(* IEC 61131-3 sources: plc-st-coding-agent/progress/evidence/f14_v10_full_20261113/jobs/codex_deepseek-v4pro, 82 files *)

(* ---- public-easy-01.candidate_01.st ---- *)
FUNCTION_BLOCK AutomatedFillingLineControl
(* ENGINEERING_CONTRACT
Stage0 idle: all outputs OFF; bottleSensor activates Pump_Motor (PUB001).
Pump_Motor: holds until cleaningConfirm; off by cleaningConfirm (PUB002).
Filling_Valve: set by cleaningConfirm; holds until fillingConfirm; off by fillingConfirm (PUB003).
Capping_Machine: set by fillingConfirm; holds until cappingConfirm; off by cappingConfirm (PUB004).
Packing_Machine: set by cappingConfirm; holds until packingConfirm; off by packingConfirm (PUB005).
Completion_Light: set by packingConfirm; holds until finishedButton; off by finishedButton (PUB006).
Same-scan priority: process only current stage trigger; at most one stage advance per scan.
Units/boundaries: BOOL outputs, integer stage 0..5; no timer or delay used.
*)
(* CONTRACT_RULES [
{"kind":"hold_until_reset","output":"Pump_Motor","set_input":"bottleSensor","reset_input":"cleaningConfirmButton"},
{"kind":"hold_until_reset","output":"Filling_Valve","set_input":"cleaningConfirmButton","reset_input":"fillingConfirmButton"},
{"kind":"hold_until_reset","output":"Capping_Machine","set_input":"fillingConfirmButton","reset_input":"cappingConfirmButton"},
{"kind":"hold_until_reset","output":"Packing_Machine","set_input":"cappingConfirmButton","reset_input":"packingConfirmButton"},
{"kind":"hold_until_reset","output":"Completion_Light","set_input":"packingConfirmButton","reset_input":"finishedButton"}
] *)
VAR_INPUT
    bottleSensor : BOOL;
    cleaningConfirmButton : BOOL;
    fillingConfirmButton : BOOL;
    cappingConfirmButton : BOOL;
    packingConfirmButton : BOOL;
    finishedButton : BOOL;
END_VAR
VAR_OUTPUT
    Pump_Motor : BOOL;
    Filling_Valve : BOOL;
    Capping_Machine : BOOL;
    Packing_Machine : BOOL;
    Completion_Light : BOOL;
END_VAR
VAR
    tmp_Stage : INT := 0;
END_VAR

IF tmp_Stage = 0 THEN
    IF bottleSensor THEN
        tmp_Stage := 1;
    END_IF;
ELSIF tmp_Stage = 1 THEN
    IF cleaningConfirmButton THEN
        tmp_Stage := 2;
    END_IF;
ELSIF tmp_Stage = 2 THEN
    IF fillingConfirmButton THEN
        tmp_Stage := 3;
    END_IF;
ELSIF tmp_Stage = 3 THEN
    IF cappingConfirmButton THEN
        tmp_Stage := 4;
    END_IF;
ELSIF tmp_Stage = 4 THEN
    IF packingConfirmButton THEN
        tmp_Stage := 5;
    END_IF;
ELSIF tmp_Stage = 5 THEN
    IF finishedButton THEN
        tmp_Stage := 0;
    END_IF;
END_IF;

Pump_Motor := (tmp_Stage = 1);
Filling_Valve := (tmp_Stage = 2);
Capping_Machine := (tmp_Stage = 3);
Packing_Machine := (tmp_Stage = 4);
Completion_Light := (tmp_Stage = 5);

END_FUNCTION_BLOCK

(* ---- public-easy-01.candidate_02.st ---- *)
FUNCTION_BLOCK AutomatedFillingLineControl
(* ENGINEERING_CONTRACT
Stage0 idle: all outputs OFF; bottleSensor activates Pump_Motor (PUB001).
Pump_Motor: holds until cleaningConfirm; off by cleaningConfirm (PUB002).
Filling_Valve: set by cleaningConfirm; holds until fillingConfirm; off by fillingConfirm (PUB003).
Capping_Machine: set by fillingConfirm; holds until cappingConfirm; off by cappingConfirm (PUB004).
Packing_Machine: set by cappingConfirm; holds until packingConfirm; off by packingConfirm (PUB005).
Completion_Light: set by packingConfirm; holds until finishedButton; off by finishedButton (PUB006).
Same-scan priority: process only current stage trigger; at most one stage advance per scan.
Units/boundaries: BOOL outputs, integer stage 0..5; no timer or delay used.
*)
(* CONTRACT_RULES [] *)
VAR_INPUT
    bottleSensor : BOOL;
    cleaningConfirmButton : BOOL;
    fillingConfirmButton : BOOL;
    cappingConfirmButton : BOOL;
    packingConfirmButton : BOOL;
    finishedButton : BOOL;
END_VAR
VAR_OUTPUT
    Pump_Motor : BOOL;
    Filling_Valve : BOOL;
    Capping_Machine : BOOL;
    Packing_Machine : BOOL;
    Completion_Light : BOOL;
END_VAR
VAR
    tmp_Stage : INT := 0;
END_VAR

IF tmp_Stage = 0 THEN
    IF bottleSensor THEN
        tmp_Stage := 1;
    END_IF;
ELSIF tmp_Stage = 1 THEN
    IF cleaningConfirmButton THEN
        tmp_Stage := 2;
    END_IF;
ELSIF tmp_Stage = 2 THEN
    IF fillingConfirmButton THEN
        tmp_Stage := 3;
    END_IF;
ELSIF tmp_Stage = 3 THEN
    IF cappingConfirmButton THEN
        tmp_Stage := 4;
    END_IF;
ELSIF tmp_Stage = 4 THEN
    IF packingConfirmButton THEN
        tmp_Stage := 5;
    END_IF;
ELSIF tmp_Stage = 5 THEN
    IF finishedButton THEN
        tmp_Stage := 0;
    END_IF;
END_IF;

Pump_Motor := (tmp_Stage = 1);
Filling_Valve := (tmp_Stage = 2);
Capping_Machine := (tmp_Stage = 3);
Packing_Machine := (tmp_Stage = 4);
Completion_Light := (tmp_Stage = 5);

END_FUNCTION_BLOCK

(* ---- public-easy-01.raw_candidate_01.st ---- *)
FUNCTION_BLOCK AutomatedFillingLineControl
(* ENGINEERING_CONTRACT
Stage0 idle: all outputs OFF; bottleSensor activates Pump_Motor (PUB001).
Pump_Motor: holds until cleaningConfirm; off by cleaningConfirm (PUB002).
Filling_Valve: set by cleaningConfirm; holds until fillingConfirm; off by fillingConfirm (PUB003).
Capping_Machine: set by fillingConfirm; holds until cappingConfirm; off by cappingConfirm (PUB004).
Packing_Machine: set by cappingConfirm; holds until packingConfirm; off by packingConfirm (PUB005).
Completion_Light: set by packingConfirm; holds until finishedButton; off by finishedButton (PUB006).
Same-scan priority: process only current stage trigger; at most one stage advance per scan.
Units/boundaries: BOOL outputs, integer stage 0..5; no timer or delay used.
*)
(* CONTRACT_RULES [
{"kind":"hold_until_reset","output":"Pump_Motor","set_input":"bottleSensor","reset_input":"cleaningConfirmButton"},
{"kind":"hold_until_reset","output":"Filling_Valve","set_input":"cleaningConfirmButton","reset_input":"fillingConfirmButton"},
{"kind":"hold_until_reset","output":"Capping_Machine","set_input":"fillingConfirmButton","reset_input":"cappingConfirmButton"},
{"kind":"hold_until_reset","output":"Packing_Machine","set_input":"cappingConfirmButton","reset_input":"packingConfirmButton"},
{"kind":"hold_until_reset","output":"Completion_Light","set_input":"packingConfirmButton","reset_input":"finishedButton"}
] *)
VAR_INPUT
    bottleSensor : BOOL;
    cleaningConfirmButton : BOOL;
    fillingConfirmButton : BOOL;
    cappingConfirmButton : BOOL;
    packingConfirmButton : BOOL;
    finishedButton : BOOL;
END_VAR
VAR_OUTPUT
    Pump_Motor : BOOL;
    Filling_Valve : BOOL;
    Capping_Machine : BOOL;
    Packing_Machine : BOOL;
    Completion_Light : BOOL;
END_VAR
VAR
    tmp_Stage : INT := 0;
END_VAR

IF tmp_Stage = 0 THEN
    IF bottleSensor THEN
        tmp_Stage := 1;
    END_IF;
ELSIF tmp_Stage = 1 THEN
    IF cleaningConfirmButton THEN
        tmp_Stage := 2;
    END_IF;
ELSIF tmp_Stage = 2 THEN
    IF fillingConfirmButton THEN
        tmp_Stage := 3;
    END_IF;
ELSIF tmp_Stage = 3 THEN
    IF cappingConfirmButton THEN
        tmp_Stage := 4;
    END_IF;
ELSIF tmp_Stage = 4 THEN
    IF packingConfirmButton THEN
        tmp_Stage := 5;
    END_IF;
ELSIF tmp_Stage = 5 THEN
    IF finishedButton THEN
        tmp_Stage := 0;
    END_IF;
END_IF;

Pump_Motor := (tmp_Stage = 1);
Filling_Valve := (tmp_Stage = 2);
Capping_Machine := (tmp_Stage = 3);
Packing_Machine := (tmp_Stage = 4);
Completion_Light := (tmp_Stage = 5);

END_FUNCTION_BLOCK

(* ---- public-easy-01.raw_candidate_02.st ---- *)
FUNCTION_BLOCK AutomatedFillingLineControl
(* ENGINEERING_CONTRACT
Stage0 idle: all outputs OFF; bottleSensor activates Pump_Motor (PUB001).
Pump_Motor: holds until cleaningConfirm; off by cleaningConfirm (PUB002).
Filling_Valve: set by cleaningConfirm; holds until fillingConfirm; off by fillingConfirm (PUB003).
Capping_Machine: set by fillingConfirm; holds until cappingConfirm; off by cappingConfirm (PUB004).
Packing_Machine: set by cappingConfirm; holds until packingConfirm; off by packingConfirm (PUB005).
Completion_Light: set by packingConfirm; holds until finishedButton; off by finishedButton (PUB006).
Same-scan priority: process only current stage trigger; at most one stage advance per scan.
Units/boundaries: BOOL outputs, integer stage 0..5; no timer or delay used.
*)
(* CONTRACT_RULES [] *)
VAR_INPUT
    bottleSensor : BOOL;
    cleaningConfirmButton : BOOL;
    fillingConfirmButton : BOOL;
    cappingConfirmButton : BOOL;
    packingConfirmButton : BOOL;
    finishedButton : BOOL;
END_VAR
VAR_OUTPUT
    Pump_Motor : BOOL;
    Filling_Valve : BOOL;
    Capping_Machine : BOOL;
    Packing_Machine : BOOL;
    Completion_Light : BOOL;
END_VAR
VAR
    tmp_Stage : INT := 0;
END_VAR

IF tmp_Stage = 0 THEN
    IF bottleSensor THEN
        tmp_Stage := 1;
    END_IF;
ELSIF tmp_Stage = 1 THEN
    IF cleaningConfirmButton THEN
        tmp_Stage := 2;
    END_IF;
ELSIF tmp_Stage = 2 THEN
    IF fillingConfirmButton THEN
        tmp_Stage := 3;
    END_IF;
ELSIF tmp_Stage = 3 THEN
    IF cappingConfirmButton THEN
        tmp_Stage := 4;
    END_IF;
ELSIF tmp_Stage = 4 THEN
    IF packingConfirmButton THEN
        tmp_Stage := 5;
    END_IF;
ELSIF tmp_Stage = 5 THEN
    IF finishedButton THEN
        tmp_Stage := 0;
    END_IF;
END_IF;

Pump_Motor := (tmp_Stage = 1);
Filling_Valve := (tmp_Stage = 2);
Capping_Machine := (tmp_Stage = 3);
Packing_Machine := (tmp_Stage = 4);
Completion_Light := (tmp_Stage = 5);

END_FUNCTION_BLOCK

(* ---- public-easy-02.candidate_01.st ---- *)
FUNCTION_BLOCK FB
(* ENGINEERING_CONTRACT
- PUB001: per-cycle edge detection on all 32 bits of DWORD value.
- hasChanged: on when current value <> retained lastValue; off otherwise.
- risingBits[i]: on when lastValue[i]=0 and value[i]=1; noOfRisingBits counts bits 0..31.
- hasRisingEdges: on when noOfRisingBits > 0; off otherwise.
- fallingBits[i]: on when lastValue[i]=1 and value[i]=0; noOfFallingBits counts bits 0..31.
- hasFallingEdges: on when noOfFallingBits > 0; off otherwise.
- Retention: only lastValue is retained. Outputs are recomputed every scan; no user reset.
- First-scan baseline: lastValue=0; unspecified, tested consistently with previous value zero.
- Priority: compare against old lastValue first, then store current value at scan end.
- Bounds: counts are USINT 0..32; masks cover DWORD bits 0..31.
*)
(* CONTRACT_RULES [] *)
VAR_INPUT
    value : DWORD;
END_VAR
VAR_OUTPUT
    hasChanged : BOOL;
    hasRisingEdges : BOOL;
    risingBits : DWORD;
    noOfRisingBits : USINT;
    hasFallingEdges : BOOL;
    fallingBits : DWORD;
    noOfFallingBits : USINT;
END_VAR
VAR
    lastValue : DWORD;
    tmp_rising : DWORD;
    tmp_falling : DWORD;
    tmp_i : INT;
END_VAR

tmp_rising := (NOT lastValue) AND value;
tmp_falling := lastValue AND (NOT value);

hasChanged := value <> lastValue;
risingBits := tmp_rising;
fallingBits := tmp_falling;

noOfRisingBits := 0;
noOfFallingBits := 0;

FOR tmp_i := 0 TO 31 DO
    IF (tmp_rising AND SHL(DWORD#1, tmp_i)) <> DWORD#0 THEN
        noOfRisingBits := noOfRisingBits + 1;
    END_IF;
    IF (tmp_falling AND SHL(DWORD#1, tmp_i)) <> DWORD#0 THEN
        noOfFallingBits := noOfFallingBits + 1;
    END_IF;
END_FOR;

hasRisingEdges := noOfRisingBits > 0;
hasFallingEdges := noOfFallingBits > 0;

lastValue := value;
END_FUNCTION_BLOCK

(* ---- public-easy-02.raw_candidate_01.st ---- *)
FUNCTION_BLOCK FB
(* ENGINEERING_CONTRACT
- PUB001: per-cycle edge detection on all 32 bits of DWORD value.
- hasChanged: on when current value <> retained lastValue; off otherwise.
- risingBits[i]: on when lastValue[i]=0 and value[i]=1; noOfRisingBits counts bits 0..31.
- hasRisingEdges: on when noOfRisingBits > 0; off otherwise.
- fallingBits[i]: on when lastValue[i]=1 and value[i]=0; noOfFallingBits counts bits 0..31.
- hasFallingEdges: on when noOfFallingBits > 0; off otherwise.
- Retention: only lastValue is retained. Outputs are recomputed every scan; no user reset.
- First-scan baseline: lastValue=0; unspecified, tested consistently with previous value zero.
- Priority: compare against old lastValue first, then store current value at scan end.
- Bounds: counts are USINT 0..32; masks cover DWORD bits 0..31.
*)
(* CONTRACT_RULES [] *)
VAR_INPUT
    value : DWORD;
END_VAR
VAR_OUTPUT
    hasChanged : BOOL;
    hasRisingEdges : BOOL;
    risingBits : DWORD;
    noOfRisingBits : USINT;
    hasFallingEdges : BOOL;
    fallingBits : DWORD;
    noOfFallingBits : USINT;
END_VAR
VAR
    lastValue : DWORD;
    tmp_rising : DWORD;
    tmp_falling : DWORD;
    tmp_i : INT;
END_VAR

tmp_rising := (NOT lastValue) AND value;
tmp_falling := lastValue AND (NOT value);

hasChanged := value <> lastValue;
risingBits := tmp_rising;
fallingBits := tmp_falling;

noOfRisingBits := 0;
noOfFallingBits := 0;

FOR tmp_i := 0 TO 31 DO
    IF (tmp_rising AND SHL(DWORD#1, tmp_i)) <> DWORD#0 THEN
        noOfRisingBits := noOfRisingBits + 1;
    END_IF;
    IF (tmp_falling AND SHL(DWORD#1, tmp_i)) <> DWORD#0 THEN
        noOfFallingBits := noOfFallingBits + 1;
    END_IF;
END_FOR;

hasRisingEdges := noOfRisingBits > 0;
hasFallingEdges := noOfFallingBits > 0;

lastValue := value;
END_FUNCTION_BLOCK

(* ---- public-easy-03.candidate_01.st ---- *)
FUNCTION_BLOCK AlarmHandling
(* ENGINEERING_CONTRACT
  hiAlarm (PUB001): activate only when Value > hiLevel; hold across deadband until deactivation.
  hiAlarm deactivation (PUB001): deactivate only when Value < hiLevel - hystWindow (strict).
  loAlarm (PUB001): activate only when Value < loLevel; hold across deadband until deactivation.
  loAlarm deactivation (PUB001): deactivate only when Value > loLevel + hystWindow (strict).
  error/status (PUB006, PUB007): normal scan sets error:=FALSE and status:=0.
  Same-scan priority: loLevel >= hiLevel (16#8001) is checked first and invokes RETURN before alarm evaluation.
  hystWindow >= hiLevel - loLevel (16#8002) is checked next and suppresses normal alarm evaluation via ELSE.
  Retention: alarm outputs persist while inside their respective hysteresis deadband.
  Units: REAL values are dimensionless; status is a hexadecimal WORD code.
  Unspecified: behavior for NaN/Inf, negative hystWindow, and historical alarm state during error scans.
*)
(* CONTRACT_RULES [] *)
VAR_INPUT
    Value      : REAL;
    hiLevel    : REAL;
    loLevel    : REAL;
    hystWindow : REAL;
END_VAR
VAR_OUTPUT
    hiAlarm : BOOL;
    loAlarm : BOOL;
    error   : BOOL;
    status  : WORD;
END_VAR
VAR
END_VAR

    error := FALSE;
    status := 0;

    IF loLevel >= hiLevel THEN
        error := TRUE;
        status := WORD#16#8001;
        RETURN;
    END_IF;

    IF hystWindow >= (hiLevel - loLevel) THEN
        error := TRUE;
        status := WORD#16#8002;
    ELSE
        IF Value > hiLevel THEN
            hiAlarm := TRUE;
        ELSIF Value < (hiLevel - hystWindow) THEN
            hiAlarm := FALSE;
        END_IF;

        IF Value < loLevel THEN
            loAlarm := TRUE;
        ELSIF Value > (loLevel + hystWindow) THEN
            loAlarm := FALSE;
        END_IF;
    END_IF;

END_FUNCTION_BLOCK

(* ---- public-easy-03.raw_candidate_01.st ---- *)
FUNCTION_BLOCK AlarmHandling
(* ENGINEERING_CONTRACT
  hiAlarm (PUB001): activate only when Value > hiLevel; hold across deadband until deactivation.
  hiAlarm deactivation (PUB001): deactivate only when Value < hiLevel - hystWindow (strict).
  loAlarm (PUB001): activate only when Value < loLevel; hold across deadband until deactivation.
  loAlarm deactivation (PUB001): deactivate only when Value > loLevel + hystWindow (strict).
  error/status (PUB006, PUB007): normal scan sets error:=FALSE and status:=0.
  Same-scan priority: loLevel >= hiLevel (16#8001) is checked first and invokes RETURN before alarm evaluation.
  hystWindow >= hiLevel - loLevel (16#8002) is checked next and suppresses normal alarm evaluation via ELSE.
  Retention: alarm outputs persist while inside their respective hysteresis deadband.
  Units: REAL values are dimensionless; status is a hexadecimal WORD code.
  Unspecified: behavior for NaN/Inf, negative hystWindow, and historical alarm state during error scans.
*)
(* CONTRACT_RULES [] *)
VAR_INPUT
    Value      : REAL;
    hiLevel    : REAL;
    loLevel    : REAL;
    hystWindow : REAL;
END_VAR
VAR_OUTPUT
    hiAlarm : BOOL;
    loAlarm : BOOL;
    error   : BOOL;
    status  : WORD;
END_VAR
VAR
END_VAR

    error := FALSE;
    status := 0;

    IF loLevel >= hiLevel THEN
        error := TRUE;
        status := WORD#16#8001;
        RETURN;
    END_IF;

    IF hystWindow >= (hiLevel - loLevel) THEN
        error := TRUE;
        status := WORD#16#8002;
    ELSE
        IF Value > hiLevel THEN
            hiAlarm := TRUE;
        ELSIF Value < (hiLevel - hystWindow) THEN
            hiAlarm := FALSE;
        END_IF;

        IF Value < loLevel THEN
            loAlarm := TRUE;
        ELSIF Value > (loLevel + hystWindow) THEN
            loAlarm := FALSE;
        END_IF;
    END_IF;

END_FUNCTION_BLOCK

(* ---- public-easy-04.candidate_01.st ---- *)
FUNCTION_BLOCK JamPumpControl
VAR_INPUT
    VISCOSITY_OK : BOOL;
    PASTE_E_STOP_NC : BOOL;
    DebounceTime : TIME;
    CycleTime : TIME;
END_VAR
VAR_OUTPUT
    VFD_RUN : BOOL := FALSE;
    PUMP_MAINT_DUE : BOOL := FALSE;
    PUMP_RUNTIME_ACC : LTIME := LTIME#0s;
END_VAR
VAR
    viscosityValid : BOOL := FALSE;
    viscosityDebounce : TON;
END_VAR

(* ENGINEERING_CONTRACT
Viscosity state PUB001/PUB002: activation after VISCOSITY_OK remains TRUE for DebounceTime via TON; invalidated immediately on VISCOSITY_OK FALSE; already-valid state retained through E-stop; incomplete debounce timing cleared on E-stop FALSE.
VFD_RUN PUB002/PUB005: activation = PASTE_E_STOP_NC AND viscosityValid; no hold/latch; E-stop FALSE disables run immediately in same scan; initialized FALSE.
PUMP_RUNTIME_ACC PUB003/PUB005: activation after current VFD_RUN computation; adds TIME_TO_LTIME(CycleTime) while VFD_RUN TRUE; retained while stopped; no explicit reset; initialized LTIME#0s.
PUMP_MAINT_DUE PUB004/PUB005: activation and retention when PUMP_RUNTIME_ACC >= LTIME#500h; no reset; informational only, never gates run/permissive; initialized FALSE.
Same-scan priority: E-stop disable and viscosity invalidation occur before run accumulation; maintenance computation is independent.
Units/boundaries: DebounceTime TIME ms, CycleTime TIME ms, PUMP_RUNTIME_ACC LTIME ns, maintenance threshold >= 500 h.
*)

(* CONTRACT_RULES [] *)

viscosityDebounce(IN := VISCOSITY_OK AND PASTE_E_STOP_NC,
                  PT := DebounceTime);

IF NOT VISCOSITY_OK THEN
    viscosityValid := FALSE;
ELSIF viscosityDebounce.Q THEN
    viscosityValid := TRUE;
END_IF;

VFD_RUN := PASTE_E_STOP_NC AND viscosityValid;

IF VFD_RUN THEN
    PUMP_RUNTIME_ACC := PUMP_RUNTIME_ACC + TIME_TO_LTIME(CycleTime);
END_IF;

IF PUMP_RUNTIME_ACC >= LTIME#500h THEN
    PUMP_MAINT_DUE := TRUE;
END_IF;

END_FUNCTION_BLOCK

(* ---- public-easy-04.raw_candidate_01.st ---- *)
FUNCTION_BLOCK JamPumpControl
VAR_INPUT
    VISCOSITY_OK : BOOL;
    PASTE_E_STOP_NC : BOOL;
    DebounceTime : TIME;
    CycleTime : TIME;
END_VAR
VAR_OUTPUT
    VFD_RUN : BOOL := FALSE;
    PUMP_MAINT_DUE : BOOL := FALSE;
    PUMP_RUNTIME_ACC : LTIME := LTIME#0s;
END_VAR
VAR
    viscosityValid : BOOL := FALSE;
    viscosityDebounce : TON;
END_VAR

(* ENGINEERING_CONTRACT
Viscosity state PUB001/PUB002: activation after VISCOSITY_OK remains TRUE for DebounceTime via TON; invalidated immediately on VISCOSITY_OK FALSE; already-valid state retained through E-stop; incomplete debounce timing cleared on E-stop FALSE.
VFD_RUN PUB002/PUB005: activation = PASTE_E_STOP_NC AND viscosityValid; no hold/latch; E-stop FALSE disables run immediately in same scan; initialized FALSE.
PUMP_RUNTIME_ACC PUB003/PUB005: activation after current VFD_RUN computation; adds TIME_TO_LTIME(CycleTime) while VFD_RUN TRUE; retained while stopped; no explicit reset; initialized LTIME#0s.
PUMP_MAINT_DUE PUB004/PUB005: activation and retention when PUMP_RUNTIME_ACC >= LTIME#500h; no reset; informational only, never gates run/permissive; initialized FALSE.
Same-scan priority: E-stop disable and viscosity invalidation occur before run accumulation; maintenance computation is independent.
Units/boundaries: DebounceTime TIME ms, CycleTime TIME ms, PUMP_RUNTIME_ACC LTIME ns, maintenance threshold >= 500 h.
*)

(* CONTRACT_RULES [] *)

viscosityDebounce(IN := VISCOSITY_OK AND PASTE_E_STOP_NC,
                  PT := DebounceTime);

IF NOT VISCOSITY_OK THEN
    viscosityValid := FALSE;
ELSIF viscosityDebounce.Q THEN
    viscosityValid := TRUE;
END_IF;

VFD_RUN := PASTE_E_STOP_NC AND viscosityValid;

IF VFD_RUN THEN
    PUMP_RUNTIME_ACC := PUMP_RUNTIME_ACC + TIME_TO_LTIME(CycleTime);
END_IF;

IF PUMP_RUNTIME_ACC >= LTIME#500h THEN
    PUMP_MAINT_DUE := TRUE;
END_IF;

END_FUNCTION_BLOCK

(* ---- public-easy-05.candidate_01.st ---- *)
FUNCTION_BLOCK WeldGapAlarmFB
VAR_INPUT
    Gap_Exceeded        : BOOL;
    Weld_E_Stop_NC      : BOOL;
    DebounceTime        : TIME;
END_VAR
VAR_OUTPUT
    Operator_Alert       : BOOL;
    Weld_Soft_Start_Active : BOOL;
END_VAR
VAR
    InitTimer       : TON;
    DebounceTimer   : TON;
    InitComplete    : BOOL;
    NormalMonitor   : BOOL;
END_VAR

(*
ENGINEERING_CONTRACT
- Operator_Alert: activates only when initialization is complete, E-stop is inactive,
  and Gap_Exceeded has remained TRUE for DebounceTime (PUB003, PUB004).
  It is FALSE during the 5 s initialization period (PUB002).
- Operator_Alert reset: immediately FALSE when Gap_Exceeded becomes FALSE or E-stop
  becomes active; normal-monitoring conditions must remain true to hold it (PUB003, PUB004).
- Debounce timing: accumulates only during initialized normal monitoring with E-stop
  inactive and resets when Gap_Exceeded is FALSE or E-stop is active (PUB002, PUB003, PUB004).
- Weld_Soft_Start_Active: TRUE only during the first 5 s after power-up, independent of
  E-stop state; it is not a speed ramp (PUB002, PUB005). E-stop state is not specified
  for this output.
- Boundaries/units: initialization is fixed T#5S; DebounceTime uses TIME milliseconds.
  TON activation occurs at elapsed time >= PT.
*)

InitTimer(IN := TRUE, PT := T#5S);
InitComplete := InitTimer.Q;
NormalMonitor := InitComplete AND Weld_E_Stop_NC;

DebounceTimer(IN := Gap_Exceeded AND NormalMonitor, PT := DebounceTime);

Operator_Alert := NormalMonitor AND DebounceTimer.Q;
Weld_Soft_Start_Active := NOT InitComplete;

(* CONTRACT_RULES [] *)
END_FUNCTION_BLOCK

(* ---- public-easy-05.raw_candidate_01.st ---- *)
FUNCTION_BLOCK WeldGapAlarmFB
VAR_INPUT
    Gap_Exceeded        : BOOL;
    Weld_E_Stop_NC      : BOOL;
    DebounceTime        : TIME;
END_VAR
VAR_OUTPUT
    Operator_Alert       : BOOL;
    Weld_Soft_Start_Active : BOOL;
END_VAR
VAR
    InitTimer       : TON;
    DebounceTimer   : TON;
    InitComplete    : BOOL;
    NormalMonitor   : BOOL;
END_VAR

(*
ENGINEERING_CONTRACT
- Operator_Alert: activates only when initialization is complete, E-stop is inactive,
  and Gap_Exceeded has remained TRUE for DebounceTime (PUB003, PUB004).
  It is FALSE during the 5 s initialization period (PUB002).
- Operator_Alert reset: immediately FALSE when Gap_Exceeded becomes FALSE or E-stop
  becomes active; normal-monitoring conditions must remain true to hold it (PUB003, PUB004).
- Debounce timing: accumulates only during initialized normal monitoring with E-stop
  inactive and resets when Gap_Exceeded is FALSE or E-stop is active (PUB002, PUB003, PUB004).
- Weld_Soft_Start_Active: TRUE only during the first 5 s after power-up, independent of
  E-stop state; it is not a speed ramp (PUB002, PUB005). E-stop state is not specified
  for this output.
- Boundaries/units: initialization is fixed T#5S; DebounceTime uses TIME milliseconds.
  TON activation occurs at elapsed time >= PT.
*)

InitTimer(IN := TRUE, PT := T#5S);
InitComplete := InitTimer.Q;
NormalMonitor := InitComplete AND Weld_E_Stop_NC;

DebounceTimer(IN := Gap_Exceeded AND NormalMonitor, PT := DebounceTime);

Operator_Alert := NormalMonitor AND DebounceTimer.Q;
Weld_Soft_Start_Active := NOT InitComplete;

(* CONTRACT_RULES [] *)
END_FUNCTION_BLOCK

(* ---- public-easy-06.candidate_01.st ---- *)
FUNCTION_BLOCK AerationBlowerDelayedStart
VAR_INPUT
    DO_LOW : BOOL;
    AERATION_E_STOP_NC : BOOL;
END_VAR
VAR_OUTPUT
    BLOWER_RUN : BOOL;
    AERATION_BLOWER_CYCLE_COUNT : UINT;
END_VAR
VAR
    tmp_StartDelay : TON;
    tmp_PrevRun : BOOL := FALSE;
END_VAR

(*
ENGINEERING_CONTRACT
- BLOWER_RUN activation: only when DO_LOW and AERATION_E_STOP_NC have both been TRUE for T#5s (PUB001).
- BLOWER_RUN retention/hold: remains TRUE only while both enabling conditions remain TRUE; no separate latch is used.
- BLOWER_RUN explicit reset/deactivation: any FALSE of DO_LOW or AERATION_E_STOP_NC clears timer IN immediately, so output and timing reset (PUB002).
- AERATION_BLOWER_CYCLE_COUNT activation: increments once on each BLOWER_RUN FALSE->TRUE transition; not repeated during continuous run (PUB003).
- AERATION_BLOWER_CYCLE_COUNT reset: initialized to zero at power-up; no task-specified runtime reset is implemented (PUB004).
- Same-scan priority: current DO_LOW/E_STOP condition directly gates TON.IN before timer Q and edge counting are evaluated.
- Units/boundaries: delay is 5 000 ms (T#5s); cycle count is UINT and unspecified at maximum rollover.
*)
(* CONTRACT_RULES [] *)

tmp_StartDelay(IN := DO_LOW AND AERATION_E_STOP_NC, PT := T#5S);

BLOWER_RUN := tmp_StartDelay.Q;

IF BLOWER_RUN AND NOT tmp_PrevRun THEN
    AERATION_BLOWER_CYCLE_COUNT := AERATION_BLOWER_CYCLE_COUNT + 1;
END_IF;

tmp_PrevRun := BLOWER_RUN;

END_FUNCTION_BLOCK

(* ---- public-easy-06.raw_candidate_01.st ---- *)
FUNCTION_BLOCK AerationBlowerDelayedStart
VAR_INPUT
    DO_LOW : BOOL;
    AERATION_E_STOP_NC : BOOL;
END_VAR
VAR_OUTPUT
    BLOWER_RUN : BOOL;
    AERATION_BLOWER_CYCLE_COUNT : UINT;
END_VAR
VAR
    tmp_StartDelay : TON;
    tmp_PrevRun : BOOL := FALSE;
END_VAR

(*
ENGINEERING_CONTRACT
- BLOWER_RUN activation: only when DO_LOW and AERATION_E_STOP_NC have both been TRUE for T#5s (PUB001).
- BLOWER_RUN retention/hold: remains TRUE only while both enabling conditions remain TRUE; no separate latch is used.
- BLOWER_RUN explicit reset/deactivation: any FALSE of DO_LOW or AERATION_E_STOP_NC clears timer IN immediately, so output and timing reset (PUB002).
- AERATION_BLOWER_CYCLE_COUNT activation: increments once on each BLOWER_RUN FALSE->TRUE transition; not repeated during continuous run (PUB003).
- AERATION_BLOWER_CYCLE_COUNT reset: initialized to zero at power-up; no task-specified runtime reset is implemented (PUB004).
- Same-scan priority: current DO_LOW/E_STOP condition directly gates TON.IN before timer Q and edge counting are evaluated.
- Units/boundaries: delay is 5 000 ms (T#5s); cycle count is UINT and unspecified at maximum rollover.
*)
(* CONTRACT_RULES [] *)

tmp_StartDelay(IN := DO_LOW AND AERATION_E_STOP_NC, PT := T#5S);

BLOWER_RUN := tmp_StartDelay.Q;

IF BLOWER_RUN AND NOT tmp_PrevRun THEN
    AERATION_BLOWER_CYCLE_COUNT := AERATION_BLOWER_CYCLE_COUNT + 1;
END_IF;

tmp_PrevRun := BLOWER_RUN;

END_FUNCTION_BLOCK

(* ---- public-hard-02.candidate_01.st ---- *)
FUNCTION_BLOCK FlexibleProcessingControl
(* ENGINEERING_CONTRACT
   conveyorLeft  : active while moving to a lower-numbered station; deactivates when the destination sensor is detected or when final delivery to station 5 is complete. No separate reset input is specified. Same-scan arrival clears both conveyors (PUB002/PUB003/PUB005).
   conveyorRight : active while moving to a higher-numbered station; deactivates when the destination sensor is detected or when final delivery to station 5 is complete. No separate reset input is specified. Same-scan arrival clears both conveyors (PUB002/PUB003/PUB005).
   Processing wait: retained in phase after arrival at station 2, 3, or 4. The matching completion input starts the next sequence movement in the same scan it is detected (PUB002/PUB003).
   Start condition: sensor1 AND station1Start initiates processing from processSequence[1]; after transition, START is not re-evaluated until the current product cycle is finished (PUB001/PUB006).
   Boundaries: processLength is active in the range 1..8; active sequence positions are processSequence[1] through processSequence[processLength]. Stations are compared as USINT values 1..5 (PUB004/PUB006).
*)
(* CONTRACT_RULES [] *)
VAR_INPUT
    processLength : USINT;
    sensor1 : BOOL;
    sensor2 : BOOL;
    sensor3 : BOOL;
    sensor4 : BOOL;
    sensor5 : BOOL;
    station1Start : BOOL;
    station2Complete : BOOL;
    station3Complete : BOOL;
    station4Complete : BOOL;
    processSequence : ARRAY[1..8] OF USINT;
END_VAR
VAR_OUTPUT
    conveyorLeft : BOOL;
    conveyorRight : BOOL;
END_VAR
VAR
    tmp_phase : USINT := 0;
    tmp_seqIndex : USINT := 1;
    tmp_currentStation : USINT := 1;
    tmp_targetStation : USINT := 0;
    tmp_destSensor : BOOL := FALSE;
    tmp_completeSignal : BOOL := FALSE;
    tmp_activeLength : USINT := 1;
END_VAR

tmp_activeLength := processLength;
IF tmp_activeLength > 8 THEN
    tmp_activeLength := 8;
END_IF;
IF tmp_activeLength < 1 THEN
    tmp_activeLength := 1;
END_IF;

conveyorLeft := FALSE;
conveyorRight := FALSE;

IF tmp_phase = 0 THEN
    IF sensor1 AND station1Start THEN
        tmp_seqIndex := 1;
        IF tmp_seqIndex <= tmp_activeLength THEN
            tmp_targetStation := processSequence[tmp_seqIndex];
            tmp_phase := 1;
        END_IF;
    END_IF;
END_IF;

IF tmp_phase = 2 THEN
    tmp_completeSignal := FALSE;
    CASE tmp_currentStation OF
        2:
            tmp_completeSignal := station2Complete;
        3:
            tmp_completeSignal := station3Complete;
        4:
            tmp_completeSignal := station4Complete;
    ELSE
        tmp_completeSignal := FALSE;
    END_CASE;

    IF tmp_completeSignal THEN
        IF tmp_seqIndex < tmp_activeLength THEN
            tmp_seqIndex := tmp_seqIndex + 1;
            IF tmp_seqIndex <= tmp_activeLength THEN
                tmp_targetStation := processSequence[tmp_seqIndex];
                tmp_phase := 1;
            END_IF;
        END_IF;
    END_IF;
END_IF;

IF tmp_phase = 1 THEN
    IF tmp_targetStation > tmp_currentStation THEN
        conveyorRight := TRUE;
    ELSIF tmp_targetStation < tmp_currentStation THEN
        conveyorLeft := TRUE;
    END_IF;

    tmp_destSensor := FALSE;
    CASE tmp_targetStation OF
        2:
            tmp_destSensor := sensor2;
        3:
            tmp_destSensor := sensor3;
        4:
            tmp_destSensor := sensor4;
        5:
            tmp_destSensor := sensor5;
    ELSE
        tmp_destSensor := FALSE;
    END_CASE;

    IF tmp_destSensor THEN
        conveyorLeft := FALSE;
        conveyorRight := FALSE;
        tmp_currentStation := tmp_targetStation;

        IF tmp_currentStation = 5 THEN
            tmp_phase := 3;
        ELSE
            tmp_phase := 2;
        END_IF;
    END_IF;
END_IF;

END_FUNCTION_BLOCK

(* ---- public-hard-02.candidate_02.st ---- *)
FUNCTION_BLOCK FlexibleProcessingControl
(* ENGINEERING_CONTRACT
   conveyorLeft  : active while moving to a lower-numbered station; deactivates when the destination sensor is detected or when final delivery to station 5 is complete. No separate reset input is specified. Same-scan arrival clears both conveyors (PUB002/PUB003/PUB005).
   conveyorRight : active while moving to a higher-numbered station; deactivates when the destination sensor is detected or when final delivery to station 5 is complete. No separate reset input is specified. Same-scan arrival clears both conveyors (PUB002/PUB003/PUB005).
   Processing wait: retained in phase after arrival at station 2, 3, or 4. The matching completion input starts the next sequence movement in the same scan it is detected (PUB002/PUB003).
   Start condition: sensor1 AND station1Start initiates processing from processSequence[1]; after transition, START is not re-evaluated until the current product cycle is finished (PUB001/PUB006). On a new start, current station returns to 1.
   Boundaries: processLength is active in the range 1..8; active sequence positions are processSequence[1] through processSequence[processLength]. Stations are compared as USINT values 1..5 (PUB004/PUB006).
*)
(* CONTRACT_RULES [] *)
VAR_INPUT
    processLength : USINT;
    sensor1 : BOOL;
    sensor2 : BOOL;
    sensor3 : BOOL;
    sensor4 : BOOL;
    sensor5 : BOOL;
    station1Start : BOOL;
    station2Complete : BOOL;
    station3Complete : BOOL;
    station4Complete : BOOL;
    processSequence : ARRAY[1..8] OF USINT;
END_VAR
VAR_OUTPUT
    conveyorLeft : BOOL;
    conveyorRight : BOOL;
END_VAR
VAR
    tmp_phase : USINT := 0;
    tmp_seqIndex : USINT := 1;
    tmp_currentStation : USINT := 1;
    tmp_targetStation : USINT := 0;
    tmp_destSensor : BOOL := FALSE;
    tmp_completeSignal : BOOL := FALSE;
    tmp_activeLength : USINT := 1;
END_VAR

tmp_activeLength := processLength;
IF tmp_activeLength > 8 THEN
    tmp_activeLength := 8;
END_IF;
IF tmp_activeLength < 1 THEN
    tmp_activeLength := 1;
END_IF;

conveyorLeft := FALSE;
conveyorRight := FALSE;

IF tmp_phase = 0 THEN
    IF sensor1 AND station1Start THEN
        tmp_seqIndex := 1;
        tmp_currentStation := 1;
        IF tmp_seqIndex <= tmp_activeLength THEN
            tmp_targetStation := processSequence[tmp_seqIndex];
            tmp_phase := 1;
        END_IF;
    END_IF;
END_IF;

IF tmp_phase = 2 THEN
    tmp_completeSignal := FALSE;
    CASE tmp_currentStation OF
        2:
            tmp_completeSignal := station2Complete;
        3:
            tmp_completeSignal := station3Complete;
        4:
            tmp_completeSignal := station4Complete;
    ELSE
        tmp_completeSignal := FALSE;
    END_CASE;

    IF tmp_completeSignal THEN
        IF tmp_seqIndex < tmp_activeLength THEN
            tmp_seqIndex := tmp_seqIndex + 1;
            IF tmp_seqIndex <= tmp_activeLength THEN
                tmp_targetStation := processSequence[tmp_seqIndex];
                tmp_phase := 1;
            END_IF;
        END_IF;
    END_IF;
END_IF;

IF tmp_phase = 1 THEN
    IF tmp_targetStation > tmp_currentStation THEN
        conveyorRight := TRUE;
    ELSIF tmp_targetStation < tmp_currentStation THEN
        conveyorLeft := TRUE;
    END_IF;

    tmp_destSensor := FALSE;
    CASE tmp_targetStation OF
        2:
            tmp_destSensor := sensor2;
        3:
            tmp_destSensor := sensor3;
        4:
            tmp_destSensor := sensor4;
        5:
            tmp_destSensor := sensor5;
    ELSE
        tmp_destSensor := FALSE;
    END_CASE;

    IF tmp_destSensor THEN
        conveyorLeft := FALSE;
        conveyorRight := FALSE;
        tmp_currentStation := tmp_targetStation;

        IF tmp_currentStation = 5 THEN
            tmp_phase := 0;
        ELSE
            tmp_phase := 2;
        END_IF;
    END_IF;
END_IF;

END_FUNCTION_BLOCK

(* ---- public-hard-02.raw_candidate_01.st ---- *)
FUNCTION_BLOCK FlexibleProcessingControl
(* ENGINEERING_CONTRACT
   conveyorLeft  : active while moving to a lower-numbered station; deactivates when the destination sensor is detected or when final delivery to station 5 is complete. No separate reset input is specified. Same-scan arrival clears both conveyors (PUB002/PUB003/PUB005).
   conveyorRight : active while moving to a higher-numbered station; deactivates when the destination sensor is detected or when final delivery to station 5 is complete. No separate reset input is specified. Same-scan arrival clears both conveyors (PUB002/PUB003/PUB005).
   Processing wait: retained in phase after arrival at station 2, 3, or 4. The matching completion input starts the next sequence movement in the same scan it is detected (PUB002/PUB003).
   Start condition: sensor1 AND station1Start initiates processing from processSequence[1]; after transition, START is not re-evaluated until the current product cycle is finished (PUB001/PUB006).
   Boundaries: processLength is active in the range 1..8; active sequence positions are processSequence[1] through processSequence[processLength]. Stations are compared as USINT values 1..5 (PUB004/PUB006).
*)
(* CONTRACT_RULES [] *)
VAR_INPUT
    processLength : USINT;
    sensor1 : BOOL;
    sensor2 : BOOL;
    sensor3 : BOOL;
    sensor4 : BOOL;
    sensor5 : BOOL;
    station1Start : BOOL;
    station2Complete : BOOL;
    station3Complete : BOOL;
    station4Complete : BOOL;
    processSequence : ARRAY[1..8] OF USINT;
END_VAR
VAR_OUTPUT
    conveyorLeft : BOOL;
    conveyorRight : BOOL;
END_VAR
VAR
    tmp_phase : USINT := 0;
    tmp_seqIndex : USINT := 1;
    tmp_currentStation : USINT := 1;
    tmp_targetStation : USINT := 0;
    tmp_destSensor : BOOL := FALSE;
    tmp_completeSignal : BOOL := FALSE;
    tmp_activeLength : USINT := 1;
END_VAR

tmp_activeLength := processLength;
IF tmp_activeLength > 8 THEN
    tmp_activeLength := 8;
END_IF;
IF tmp_activeLength < 1 THEN
    tmp_activeLength := 1;
END_IF;

conveyorLeft := FALSE;
conveyorRight := FALSE;

IF tmp_phase = 0 THEN
    IF sensor1 AND station1Start THEN
        tmp_seqIndex := 1;
        IF tmp_seqIndex <= tmp_activeLength THEN
            tmp_targetStation := processSequence[tmp_seqIndex];
            tmp_phase := 1;
        END_IF;
    END_IF;
END_IF;

IF tmp_phase = 2 THEN
    tmp_completeSignal := FALSE;
    CASE tmp_currentStation OF
        2:
            tmp_completeSignal := station2Complete;
        3:
            tmp_completeSignal := station3Complete;
        4:
            tmp_completeSignal := station4Complete;
    ELSE
        tmp_completeSignal := FALSE;
    END_CASE;

    IF tmp_completeSignal THEN
        IF tmp_seqIndex < tmp_activeLength THEN
            tmp_seqIndex := tmp_seqIndex + 1;
            IF tmp_seqIndex <= tmp_activeLength THEN
                tmp_targetStation := processSequence[tmp_seqIndex];
                tmp_phase := 1;
            END_IF;
        END_IF;
    END_IF;
END_IF;

IF tmp_phase = 1 THEN
    IF tmp_targetStation > tmp_currentStation THEN
        conveyorRight := TRUE;
    ELSIF tmp_targetStation < tmp_currentStation THEN
        conveyorLeft := TRUE;
    END_IF;

    tmp_destSensor := FALSE;
    CASE tmp_targetStation OF
        2:
            tmp_destSensor := sensor2;
        3:
            tmp_destSensor := sensor3;
        4:
            tmp_destSensor := sensor4;
        5:
            tmp_destSensor := sensor5;
    ELSE
        tmp_destSensor := FALSE;
    END_CASE;

    IF tmp_destSensor THEN
        conveyorLeft := FALSE;
        conveyorRight := FALSE;
        tmp_currentStation := tmp_targetStation;

        IF tmp_currentStation = 5 THEN
            tmp_phase := 3;
        ELSE
            tmp_phase := 2;
        END_IF;
    END_IF;
END_IF;

END_FUNCTION_BLOCK

(* ---- public-hard-02.raw_candidate_02.st ---- *)
FUNCTION_BLOCK FlexibleProcessingControl
(* ENGINEERING_CONTRACT
   conveyorLeft  : active while moving to a lower-numbered station; deactivates when the destination sensor is detected or when final delivery to station 5 is complete. No separate reset input is specified. Same-scan arrival clears both conveyors (PUB002/PUB003/PUB005).
   conveyorRight : active while moving to a higher-numbered station; deactivates when the destination sensor is detected or when final delivery to station 5 is complete. No separate reset input is specified. Same-scan arrival clears both conveyors (PUB002/PUB003/PUB005).
   Processing wait: retained in phase after arrival at station 2, 3, or 4. The matching completion input starts the next sequence movement in the same scan it is detected (PUB002/PUB003).
   Start condition: sensor1 AND station1Start initiates processing from processSequence[1]; after transition, START is not re-evaluated until the current product cycle is finished (PUB001/PUB006). On a new start, current station returns to 1.
   Boundaries: processLength is active in the range 1..8; active sequence positions are processSequence[1] through processSequence[processLength]. Stations are compared as USINT values 1..5 (PUB004/PUB006).
*)
(* CONTRACT_RULES [] *)
VAR_INPUT
    processLength : USINT;
    sensor1 : BOOL;
    sensor2 : BOOL;
    sensor3 : BOOL;
    sensor4 : BOOL;
    sensor5 : BOOL;
    station1Start : BOOL;
    station2Complete : BOOL;
    station3Complete : BOOL;
    station4Complete : BOOL;
    processSequence : ARRAY[1..8] OF USINT;
END_VAR
VAR_OUTPUT
    conveyorLeft : BOOL;
    conveyorRight : BOOL;
END_VAR
VAR
    tmp_phase : USINT := 0;
    tmp_seqIndex : USINT := 1;
    tmp_currentStation : USINT := 1;
    tmp_targetStation : USINT := 0;
    tmp_destSensor : BOOL := FALSE;
    tmp_completeSignal : BOOL := FALSE;
    tmp_activeLength : USINT := 1;
END_VAR

tmp_activeLength := processLength;
IF tmp_activeLength > 8 THEN
    tmp_activeLength := 8;
END_IF;
IF tmp_activeLength < 1 THEN
    tmp_activeLength := 1;
END_IF;

conveyorLeft := FALSE;
conveyorRight := FALSE;

IF tmp_phase = 0 THEN
    IF sensor1 AND station1Start THEN
        tmp_seqIndex := 1;
        tmp_currentStation := 1;
        IF tmp_seqIndex <= tmp_activeLength THEN
            tmp_targetStation := processSequence[tmp_seqIndex];
            tmp_phase := 1;
        END_IF;
    END_IF;
END_IF;

IF tmp_phase = 2 THEN
    tmp_completeSignal := FALSE;
    CASE tmp_currentStation OF
        2:
            tmp_completeSignal := station2Complete;
        3:
            tmp_completeSignal := station3Complete;
        4:
            tmp_completeSignal := station4Complete;
    ELSE
        tmp_completeSignal := FALSE;
    END_CASE;

    IF tmp_completeSignal THEN
        IF tmp_seqIndex < tmp_activeLength THEN
            tmp_seqIndex := tmp_seqIndex + 1;
            IF tmp_seqIndex <= tmp_activeLength THEN
                tmp_targetStation := processSequence[tmp_seqIndex];
                tmp_phase := 1;
            END_IF;
        END_IF;
    END_IF;
END_IF;

IF tmp_phase = 1 THEN
    IF tmp_targetStation > tmp_currentStation THEN
        conveyorRight := TRUE;
    ELSIF tmp_targetStation < tmp_currentStation THEN
        conveyorLeft := TRUE;
    END_IF;

    tmp_destSensor := FALSE;
    CASE tmp_targetStation OF
        2:
            tmp_destSensor := sensor2;
        3:
            tmp_destSensor := sensor3;
        4:
            tmp_destSensor := sensor4;
        5:
            tmp_destSensor := sensor5;
    ELSE
        tmp_destSensor := FALSE;
    END_CASE;

    IF tmp_destSensor THEN
        conveyorLeft := FALSE;
        conveyorRight := FALSE;
        tmp_currentStation := tmp_targetStation;

        IF tmp_currentStation = 5 THEN
            tmp_phase := 0;
        ELSE
            tmp_phase := 2;
        END_IF;
    END_IF;
END_IF;

END_FUNCTION_BLOCK

(* ---- public-hard-03.candidate_01.st ---- *)
TYPE ST_Recipe :
STRUCT
    recipeID : INT;
    ingredientType : INT;
    ingredientRatio : REAL;
    productionTemperature : REAL;
END_STRUCT
END_TYPE;

(* ENGINEERING_CONTRACT
   Outputs: success flags are same-scan level, not latched; they deactivate on the next scan (PUB003-PUB005).
   recipeQueryResult: updated only for a successful query; otherwise zeroed each scan (PUB002).
   error/status: cleared at scan start; first operation error in the scan retains error and code (PUB002-PUB005).
   Add: duplicate check before empty-slot check; uses first empty index; whole struct copy (PUB003).
   Delete: nonzero-ID match; sets only recipeID to 0 (PUB004).
   Modify: nonzero-ID match; whole struct replacement (PUB005).
   Query: nonzero-ID match; whole struct copy to result; missing ID gives 16#8001 (PUB002).
   Array bounds: 1..10; recipeID=0 denotes unused slot and is never returned as a stored recipe.
   Multiple requests: unspecified; processed add/delete/modify/query in interface order on evolving database.
*)
(* CONTRACT_RULES [] *)

FUNCTION_BLOCK RecipeManagementSystem
VAR_INPUT
    addRecipe : BOOL;
    deleteRecipe : BOOL;
    modifyRecipe : BOOL;
    queryRecipe : BOOL;
    recipeIn : ST_Recipe;
END_VAR
VAR_OUTPUT
    recipeAdded : BOOL;
    recipeDeleted : BOOL;
    recipeModified : BOOL;
    recipeQueryResult : ST_Recipe;
    error : BOOL;
    status : WORD;
END_VAR
VAR_IN_OUT
    recipe : ARRAY[1..10] OF ST_Recipe;
END_VAR
VAR
    tmp_i : INT;
    tmp_foundIndex : INT;
    tmp_emptyIndex : INT;
    tmp_found : BOOL;
END_VAR

recipeAdded := FALSE;
recipeDeleted := FALSE;
recipeModified := FALSE;
recipeQueryResult.recipeID := 0;
recipeQueryResult.ingredientType := 0;
recipeQueryResult.ingredientRatio := 0.0;
recipeQueryResult.productionTemperature := 0.0;
error := FALSE;
status := 16#0000;

IF addRecipe THEN
    tmp_found := FALSE;
    tmp_emptyIndex := 0;

    FOR tmp_i := 1 TO 10 DO
        IF recipe[tmp_i].recipeID = recipeIn.recipeID THEN
            tmp_found := TRUE;
        END_IF;

        IF (recipe[tmp_i].recipeID = 0) AND (tmp_emptyIndex = 0) THEN
            tmp_emptyIndex := tmp_i;
        END_IF;
    END_FOR;

    IF tmp_found THEN
        IF NOT error THEN
            error := TRUE;
            status := 16#8002;
        END_IF;
    ELSIF tmp_emptyIndex = 0 THEN
        IF NOT error THEN
            error := TRUE;
            status := 16#8003;
        END_IF;
    ELSE
        recipe[tmp_emptyIndex] := recipeIn;
        recipeAdded := TRUE;
    END_IF;
END_IF;

IF deleteRecipe THEN
    tmp_found := FALSE;
    tmp_foundIndex := 0;

    FOR tmp_i := 1 TO 10 DO
        IF (recipe[tmp_i].recipeID <> 0) AND
           (recipe[tmp_i].recipeID = recipeIn.recipeID) THEN
            tmp_found := TRUE;
            tmp_foundIndex := tmp_i;
        END_IF;
    END_FOR;

    IF NOT tmp_found THEN
        IF NOT error THEN
            error := TRUE;
            status := 16#8004;
        END_IF;
    ELSE
        recipe[tmp_foundIndex].recipeID := 0;
        recipeDeleted := TRUE;
    END_IF;
END_IF;

IF modifyRecipe THEN
    tmp_found := FALSE;
    tmp_foundIndex := 0;

    FOR tmp_i := 1 TO 10 DO
        IF (recipe[tmp_i].recipeID <> 0) AND
           (recipe[tmp_i].recipeID = recipeIn.recipeID) THEN
            tmp_found := TRUE;
            tmp_foundIndex := tmp_i;
        END_IF;
    END_FOR;

    IF NOT tmp_found THEN
        IF NOT error THEN
            error := TRUE;
            status := 16#8005;
        END_IF;
    ELSE
        recipe[tmp_foundIndex] := recipeIn;
        recipeModified := TRUE;
    END_IF;
END_IF;

IF queryRecipe THEN
    tmp_found := FALSE;
    tmp_foundIndex := 0;

    FOR tmp_i := 1 TO 10 DO
        IF (recipe[tmp_i].recipeID <> 0) AND
           (recipe[tmp_i].recipeID = recipeIn.recipeID) THEN
            tmp_found := TRUE;
            tmp_foundIndex := tmp_i;
        END_IF;
    END_FOR;

    IF NOT tmp_found THEN
        IF NOT error THEN
            error := TRUE;
            status := 16#8001;
        END_IF;
    ELSE
        recipeQueryResult := recipe[tmp_foundIndex];
    END_IF;
END_IF;

END_FUNCTION_BLOCK

(* ---- public-hard-03.candidate_02.st ---- *)
TYPE ST_Recipe :
STRUCT
    recipeID : INT;
    ingredientType : INT;
    ingredientRatio : REAL;
    productionTemperature : REAL;
END_STRUCT
END_TYPE;

(* ENGINEERING_CONTRACT
   Outputs: success flags are same-scan level, not latched; they deactivate on the next scan (PUB003-PUB005).
   recipeQueryResult: updated only for a successful query; otherwise zeroed each scan (PUB002).
   error/status: cleared at scan start; a reported operation error retains error and code for that invocation (PUB002-PUB005).
   Add: duplicate check before empty-slot check; uses first empty index; whole struct copy (PUB003).
   Delete: nonzero-ID match; sets only recipeID to 0 (PUB004).
   Modify: nonzero-ID match; whole struct replacement (PUB005).
   Query: nonzero-ID match; whole struct copy to result; missing ID gives 16#8001 (PUB002).
   Array bounds: 1..10; recipeID=0 denotes unused slot and is never returned as a stored recipe.
   Multiple requests: unspecified by the public contract. They are reported as an unsupported combination with
   error=TRUE, status=16#8000, no database update, no success flag, and no query result.
*)
(* CONTRACT_RULES [] *)

FUNCTION_BLOCK RecipeManagementSystem
VAR_INPUT
    addRecipe : BOOL;
    deleteRecipe : BOOL;
    modifyRecipe : BOOL;
    queryRecipe : BOOL;
    recipeIn : ST_Recipe;
END_VAR
VAR_OUTPUT
    recipeAdded : BOOL;
    recipeDeleted : BOOL;
    recipeModified : BOOL;
    recipeQueryResult : ST_Recipe;
    error : BOOL;
    status : WORD;
END_VAR
VAR_IN_OUT
    recipe : ARRAY[1..10] OF ST_Recipe;
END_VAR
VAR
    tmp_i : INT;
    tmp_foundIndex : INT;
    tmp_emptyIndex : INT;
    tmp_found : BOOL;
    tmp_cmdCount : INT;
END_VAR

recipeAdded := FALSE;
recipeDeleted := FALSE;
recipeModified := FALSE;
recipeQueryResult.recipeID := 0;
recipeQueryResult.ingredientType := 0;
recipeQueryResult.ingredientRatio := 0.0;
recipeQueryResult.productionTemperature := 0.0;
error := FALSE;
status := 16#0000;

tmp_cmdCount := 0;
IF addRecipe THEN
    tmp_cmdCount := tmp_cmdCount + 1;
END_IF;
IF deleteRecipe THEN
    tmp_cmdCount := tmp_cmdCount + 1;
END_IF;
IF modifyRecipe THEN
    tmp_cmdCount := tmp_cmdCount + 1;
END_IF;
IF queryRecipe THEN
    tmp_cmdCount := tmp_cmdCount + 1;
END_IF;

IF tmp_cmdCount > 1 THEN
    error := TRUE;
    status := 16#8000;
ELSE
    IF addRecipe THEN
        tmp_found := FALSE;
        tmp_emptyIndex := 0;

        FOR tmp_i := 1 TO 10 DO
            IF recipe[tmp_i].recipeID = recipeIn.recipeID THEN
                tmp_found := TRUE;
            END_IF;

            IF (recipe[tmp_i].recipeID = 0) AND (tmp_emptyIndex = 0) THEN
                tmp_emptyIndex := tmp_i;
            END_IF;
        END_FOR;

        IF tmp_found THEN
            IF NOT error THEN
                error := TRUE;
                status := 16#8002;
            END_IF;
        ELSIF tmp_emptyIndex = 0 THEN
            IF NOT error THEN
                error := TRUE;
                status := 16#8003;
            END_IF;
        ELSE
            recipe[tmp_emptyIndex] := recipeIn;
            recipeAdded := TRUE;
        END_IF;
    END_IF;

    IF deleteRecipe THEN
        tmp_found := FALSE;
        tmp_foundIndex := 0;

        FOR tmp_i := 1 TO 10 DO
            IF (recipe[tmp_i].recipeID <> 0) AND
               (recipe[tmp_i].recipeID = recipeIn.recipeID) THEN
                tmp_found := TRUE;
                tmp_foundIndex := tmp_i;
            END_IF;
        END_FOR;

        IF NOT tmp_found THEN
            IF NOT error THEN
                error := TRUE;
                status := 16#8004;
            END_IF;
        ELSE
            recipe[tmp_foundIndex].recipeID := 0;
            recipeDeleted := TRUE;
        END_IF;
    END_IF;

    IF modifyRecipe THEN
        tmp_found := FALSE;
        tmp_foundIndex := 0;

        FOR tmp_i := 1 TO 10 DO
            IF (recipe[tmp_i].recipeID <> 0) AND
               (recipe[tmp_i].recipeID = recipeIn.recipeID) THEN
                tmp_found := TRUE;
                tmp_foundIndex := tmp_i;
            END_IF;
        END_FOR;

        IF NOT tmp_found THEN
            IF NOT error THEN
                error := TRUE;
                status := 16#8005;
            END_IF;
        ELSE
            recipe[tmp_foundIndex] := recipeIn;
            recipeModified := TRUE;
        END_IF;
    END_IF;

    IF queryRecipe THEN
        tmp_found := FALSE;
        tmp_foundIndex := 0;

        FOR tmp_i := 1 TO 10 DO
            IF (recipe[tmp_i].recipeID <> 0) AND
               (recipe[tmp_i].recipeID = recipeIn.recipeID) THEN
                tmp_found := TRUE;
                tmp_foundIndex := tmp_i;
            END_IF;
        END_FOR;

        IF NOT tmp_found THEN
            IF NOT error THEN
                error := TRUE;
                status := 16#8001;
            END_IF;
        ELSE
            recipeQueryResult := recipe[tmp_foundIndex];
        END_IF;
    END_IF;
END_IF;

END_FUNCTION_BLOCK

(* ---- public-hard-03.raw_candidate_01.st ---- *)
TYPE ST_Recipe :
STRUCT
    recipeID : INT;
    ingredientType : INT;
    ingredientRatio : REAL;
    productionTemperature : REAL;
END_STRUCT
END_TYPE

(* ENGINEERING_CONTRACT
   Outputs: success flags are same-scan level, not latched; they deactivate on the next scan (PUB003-PUB005).
   recipeQueryResult: updated only for a successful query; otherwise zeroed each scan (PUB002).
   error/status: cleared at scan start; first operation error in the scan retains error and code (PUB002-PUB005).
   Add: duplicate check before empty-slot check; uses first empty index; whole struct copy (PUB003).
   Delete: nonzero-ID match; sets only recipeID to 0 (PUB004).
   Modify: nonzero-ID match; whole struct replacement (PUB005).
   Query: nonzero-ID match; whole struct copy to result; missing ID gives 16#8001 (PUB002).
   Array bounds: 1..10; recipeID=0 denotes unused slot and is never returned as a stored recipe.
   Multiple requests: unspecified; processed add/delete/modify/query in interface order on evolving database.
*)
(* CONTRACT_RULES [] *)

FUNCTION_BLOCK RecipeManagementSystem
VAR_INPUT
    addRecipe : BOOL;
    deleteRecipe : BOOL;
    modifyRecipe : BOOL;
    queryRecipe : BOOL;
    recipeIn : ST_Recipe;
END_VAR
VAR_OUTPUT
    recipeAdded : BOOL;
    recipeDeleted : BOOL;
    recipeModified : BOOL;
    recipeQueryResult : ST_Recipe;
    error : BOOL;
    status : WORD;
END_VAR
VAR_IN_OUT
    recipe : ARRAY[1..10] OF ST_Recipe;
END_VAR
VAR
    tmp_i : INT;
    tmp_foundIndex : INT;
    tmp_emptyIndex : INT;
    tmp_found : BOOL;
END_VAR

recipeAdded := FALSE;
recipeDeleted := FALSE;
recipeModified := FALSE;
recipeQueryResult.recipeID := 0;
recipeQueryResult.ingredientType := 0;
recipeQueryResult.ingredientRatio := 0.0;
recipeQueryResult.productionTemperature := 0.0;
error := FALSE;
status := 16#0000;

IF addRecipe THEN
    tmp_found := FALSE;
    tmp_emptyIndex := 0;

    FOR tmp_i := 1 TO 10 DO
        IF recipe[tmp_i].recipeID = recipeIn.recipeID THEN
            tmp_found := TRUE;
        END_IF;

        IF (recipe[tmp_i].recipeID = 0) AND (tmp_emptyIndex = 0) THEN
            tmp_emptyIndex := tmp_i;
        END_IF;
    END_FOR;

    IF tmp_found THEN
        IF NOT error THEN
            error := TRUE;
            status := 16#8002;
        END_IF;
    ELSIF tmp_emptyIndex = 0 THEN
        IF NOT error THEN
            error := TRUE;
            status := 16#8003;
        END_IF;
    ELSE
        recipe[tmp_emptyIndex] := recipeIn;
        recipeAdded := TRUE;
    END_IF;
END_IF;

IF deleteRecipe THEN
    tmp_found := FALSE;
    tmp_foundIndex := 0;

    FOR tmp_i := 1 TO 10 DO
        IF (recipe[tmp_i].recipeID <> 0) AND
           (recipe[tmp_i].recipeID = recipeIn.recipeID) THEN
            tmp_found := TRUE;
            tmp_foundIndex := tmp_i;
        END_IF;
    END_FOR;

    IF NOT tmp_found THEN
        IF NOT error THEN
            error := TRUE;
            status := 16#8004;
        END_IF;
    ELSE
        recipe[tmp_foundIndex].recipeID := 0;
        recipeDeleted := TRUE;
    END_IF;
END_IF;

IF modifyRecipe THEN
    tmp_found := FALSE;
    tmp_foundIndex := 0;

    FOR tmp_i := 1 TO 10 DO
        IF (recipe[tmp_i].recipeID <> 0) AND
           (recipe[tmp_i].recipeID = recipeIn.recipeID) THEN
            tmp_found := TRUE;
            tmp_foundIndex := tmp_i;
        END_IF;
    END_FOR;

    IF NOT tmp_found THEN
        IF NOT error THEN
            error := TRUE;
            status := 16#8005;
        END_IF;
    ELSE
        recipe[tmp_foundIndex] := recipeIn;
        recipeModified := TRUE;
    END_IF;
END_IF;

IF queryRecipe THEN
    tmp_found := FALSE;
    tmp_foundIndex := 0;

    FOR tmp_i := 1 TO 10 DO
        IF (recipe[tmp_i].recipeID <> 0) AND
           (recipe[tmp_i].recipeID = recipeIn.recipeID) THEN
            tmp_found := TRUE;
            tmp_foundIndex := tmp_i;
        END_IF;
    END_FOR;

    IF NOT tmp_found THEN
        IF NOT error THEN
            error := TRUE;
            status := 16#8001;
        END_IF;
    ELSE
        recipeQueryResult := recipe[tmp_foundIndex];
    END_IF;
END_IF;

END_FUNCTION_BLOCK

(* ---- public-hard-03.raw_candidate_02.st ---- *)
TYPE ST_Recipe :
STRUCT
    recipeID : INT;
    ingredientType : INT;
    ingredientRatio : REAL;
    productionTemperature : REAL;
END_STRUCT
END_TYPE;

(* ENGINEERING_CONTRACT
   Outputs: success flags are same-scan level, not latched; they deactivate on the next scan (PUB003-PUB005).
   recipeQueryResult: updated only for a successful query; otherwise zeroed each scan (PUB002).
   error/status: cleared at scan start; a reported operation error retains error and code for that invocation (PUB002-PUB005).
   Add: duplicate check before empty-slot check; uses first empty index; whole struct copy (PUB003).
   Delete: nonzero-ID match; sets only recipeID to 0 (PUB004).
   Modify: nonzero-ID match; whole struct replacement (PUB005).
   Query: nonzero-ID match; whole struct copy to result; missing ID gives 16#8001 (PUB002).
   Array bounds: 1..10; recipeID=0 denotes unused slot and is never returned as a stored recipe.
   Multiple requests: unspecified by the public contract. They are reported as an unsupported combination with
   error=TRUE, status=16#8000, no database update, no success flag, and no query result.
*)
(* CONTRACT_RULES [] *)

FUNCTION_BLOCK RecipeManagementSystem
VAR_INPUT
    addRecipe : BOOL;
    deleteRecipe : BOOL;
    modifyRecipe : BOOL;
    queryRecipe : BOOL;
    recipeIn : ST_Recipe;
END_VAR
VAR_OUTPUT
    recipeAdded : BOOL;
    recipeDeleted : BOOL;
    recipeModified : BOOL;
    recipeQueryResult : ST_Recipe;
    error : BOOL;
    status : WORD;
END_VAR
VAR_IN_OUT
    recipe : ARRAY[1..10] OF ST_Recipe;
END_VAR
VAR
    tmp_i : INT;
    tmp_foundIndex : INT;
    tmp_emptyIndex : INT;
    tmp_found : BOOL;
    tmp_cmdCount : INT;
END_VAR

recipeAdded := FALSE;
recipeDeleted := FALSE;
recipeModified := FALSE;
recipeQueryResult.recipeID := 0;
recipeQueryResult.ingredientType := 0;
recipeQueryResult.ingredientRatio := 0.0;
recipeQueryResult.productionTemperature := 0.0;
error := FALSE;
status := 16#0000;

tmp_cmdCount := 0;
IF addRecipe THEN
    tmp_cmdCount := tmp_cmdCount + 1;
END_IF;
IF deleteRecipe THEN
    tmp_cmdCount := tmp_cmdCount + 1;
END_IF;
IF modifyRecipe THEN
    tmp_cmdCount := tmp_cmdCount + 1;
END_IF;
IF queryRecipe THEN
    tmp_cmdCount := tmp_cmdCount + 1;
END_IF;

IF tmp_cmdCount > 1 THEN
    error := TRUE;
    status := 16#8000;
ELSE
    IF addRecipe THEN
        tmp_found := FALSE;
        tmp_emptyIndex := 0;

        FOR tmp_i := 1 TO 10 DO
            IF recipe[tmp_i].recipeID = recipeIn.recipeID THEN
                tmp_found := TRUE;
            END_IF;

            IF (recipe[tmp_i].recipeID = 0) AND (tmp_emptyIndex = 0) THEN
                tmp_emptyIndex := tmp_i;
            END_IF;
        END_FOR;

        IF tmp_found THEN
            IF NOT error THEN
                error := TRUE;
                status := 16#8002;
            END_IF;
        ELSIF tmp_emptyIndex = 0 THEN
            IF NOT error THEN
                error := TRUE;
                status := 16#8003;
            END_IF;
        ELSE
            recipe[tmp_emptyIndex] := recipeIn;
            recipeAdded := TRUE;
        END_IF;
    END_IF;

    IF deleteRecipe THEN
        tmp_found := FALSE;
        tmp_foundIndex := 0;

        FOR tmp_i := 1 TO 10 DO
            IF (recipe[tmp_i].recipeID <> 0) AND
               (recipe[tmp_i].recipeID = recipeIn.recipeID) THEN
                tmp_found := TRUE;
                tmp_foundIndex := tmp_i;
            END_IF;
        END_FOR;

        IF NOT tmp_found THEN
            IF NOT error THEN
                error := TRUE;
                status := 16#8004;
            END_IF;
        ELSE
            recipe[tmp_foundIndex].recipeID := 0;
            recipeDeleted := TRUE;
        END_IF;
    END_IF;

    IF modifyRecipe THEN
        tmp_found := FALSE;
        tmp_foundIndex := 0;

        FOR tmp_i := 1 TO 10 DO
            IF (recipe[tmp_i].recipeID <> 0) AND
               (recipe[tmp_i].recipeID = recipeIn.recipeID) THEN
                tmp_found := TRUE;
                tmp_foundIndex := tmp_i;
            END_IF;
        END_FOR;

        IF NOT tmp_found THEN
            IF NOT error THEN
                error := TRUE;
                status := 16#8005;
            END_IF;
        ELSE
            recipe[tmp_foundIndex] := recipeIn;
            recipeModified := TRUE;
        END_IF;
    END_IF;

    IF queryRecipe THEN
        tmp_found := FALSE;
        tmp_foundIndex := 0;

        FOR tmp_i := 1 TO 10 DO
            IF (recipe[tmp_i].recipeID <> 0) AND
               (recipe[tmp_i].recipeID = recipeIn.recipeID) THEN
                tmp_found := TRUE;
                tmp_foundIndex := tmp_i;
            END_IF;
        END_FOR;

        IF NOT tmp_found THEN
            IF NOT error THEN
                error := TRUE;
                status := 16#8001;
            END_IF;
        ELSE
            recipeQueryResult := recipe[tmp_foundIndex];
        END_IF;
    END_IF;
END_IF;

END_FUNCTION_BLOCK

(* ---- public-hard-04.candidate_01.st ---- *)
FUNCTION_BLOCK FB_FIFO
VAR_INPUT
    enqueue : BOOL;
    dequeue : BOOL;
    reset : BOOL;
END_VAR
VAR_OUTPUT
    elementCount : DINT;
    status : WORD;
END_VAR
VAR_IN_OUT
    item : VARIANT;
    buffer : VARIANT;
END_VAR
VAR
    localCapacity : DINT;
    localLower : DINT;
    localHead : DINT;
    localTail : DINT;
    localCount : DINT;
    localNext : DINT;
    localLastEnqueue : BOOL;
    localLastDequeue : BOOL;
    localRisingEnqueue : BOOL;
    localRisingDequeue : BOOL;
END_VAR

(* ENGINEERING_CONTRACT
   validCount: activated by successful enqueue/dequeue; reset to 0 by reset (PUB001/PUB003).
   elementCount: mirror of persistent validCount each scan; reset sets it to 0 (PUB003/PUB004).
   status: default 16#0000; 16#8001 empty dequeue reject; 16#8002 full enqueue reject (PUB005).
   head/tail: internal only, initialized to buffer lower bound, advanced circularly (PUB006).
   priority: reset is processed before all queue operations (PUB003).
   same scan: caller precondition forbids simultaneous edges; if both occur enqueue is handled first (PUB002).
   full condition: validCount = capacity; empty condition: validCount = 0 (PUB004).
   capacity: UPPER_BOUND(buffer,1)-LOWER_BOUND(buffer,1)+1; indices are DINT (PUB004/PUB006).
   rejected operations: item and queue are not modified (PUB005).
   units/bounds: elementCount DINT 0..capacity; status WORD; no unconditional public BOOL latch.
*)

(* CONTRACT_RULES [] *)

IF localCapacity = 0 THEN
    localLower := LOWER_BOUND(buffer, 1);
    localCapacity := UPPER_BOUND(buffer, 1) - localLower + 1;
    localHead := localLower;
    localTail := localLower;
    localCount := 0;
END_IF;

status := WORD#16#0000;

localRisingEnqueue := enqueue AND NOT localLastEnqueue;
localRisingDequeue := dequeue AND NOT localLastDequeue;

IF reset THEN
    localCount := 0;
    localHead := localLower;
    localTail := localLower;
ELSE
    IF localRisingEnqueue THEN
        IF localCount < localCapacity THEN
            buffer[localTail] := item;
            localNext := localTail - localLower + 1;
            IF localNext >= localCapacity THEN
                localNext := 0;
            END_IF;
            localTail := localLower + localNext;
            localCount := localCount + 1;
        ELSE
            status := WORD#16#8002;
        END_IF;
    END_IF;

    IF localRisingDequeue THEN
        IF localCount > 0 THEN
            item := buffer[localHead];
            localNext := localHead - localLower + 1;
            IF localNext >= localCapacity THEN
                localNext := 0;
            END_IF;
            localHead := localLower + localNext;
            localCount := localCount - 1;
        ELSE
            status := WORD#16#8001;
        END_IF;
    END_IF;
END_IF;

elementCount := localCount;

localLastEnqueue := enqueue;
localLastDequeue := dequeue;

END_FUNCTION_BLOCK

(* ---- public-hard-04.raw_candidate_01.st ---- *)
FUNCTION_BLOCK FB_FIFO
VAR_INPUT
    enqueue : BOOL;
    dequeue : BOOL;
    reset : BOOL;
END_VAR
VAR_OUTPUT
    elementCount : DINT;
    status : WORD;
END_VAR
VAR_IN_OUT
    item : VARIANT;
    buffer : VARIANT;
END_VAR
VAR
    localCapacity : DINT;
    localLower : DINT;
    localHead : DINT;
    localTail : DINT;
    localCount : DINT;
    localNext : DINT;
    localLastEnqueue : BOOL;
    localLastDequeue : BOOL;
    localRisingEnqueue : BOOL;
    localRisingDequeue : BOOL;
END_VAR

(* ENGINEERING_CONTRACT
   validCount: activated by successful enqueue/dequeue; reset to 0 by reset (PUB001/PUB003).
   elementCount: mirror of persistent validCount each scan; reset sets it to 0 (PUB003/PUB004).
   status: default 16#0000; 16#8001 empty dequeue reject; 16#8002 full enqueue reject (PUB005).
   head/tail: internal only, initialized to buffer lower bound, advanced circularly (PUB006).
   priority: reset is processed before all queue operations (PUB003).
   same scan: caller precondition forbids simultaneous edges; if both occur enqueue is handled first (PUB002).
   full condition: validCount = capacity; empty condition: validCount = 0 (PUB004).
   capacity: UPPER_BOUND(buffer,1)-LOWER_BOUND(buffer,1)+1; indices are DINT (PUB004/PUB006).
   rejected operations: item and queue are not modified (PUB005).
   units/bounds: elementCount DINT 0..capacity; status WORD; no unconditional public BOOL latch.
*)

(* CONTRACT_RULES [] *)

IF localCapacity = 0 THEN
    localLower := LOWER_BOUND(buffer, 1);
    localCapacity := UPPER_BOUND(buffer, 1) - localLower + 1;
    localHead := localLower;
    localTail := localLower;
    localCount := 0;
END_IF;

status := WORD#16#0000;

localRisingEnqueue := enqueue AND NOT localLastEnqueue;
localRisingDequeue := dequeue AND NOT localLastDequeue;

IF reset THEN
    localCount := 0;
    localHead := localLower;
    localTail := localLower;
ELSE
    IF localRisingEnqueue THEN
        IF localCount < localCapacity THEN
            buffer[localTail] := item;
            localNext := localTail - localLower + 1;
            IF localNext >= localCapacity THEN
                localNext := 0;
            END_IF;
            localTail := localLower + localNext;
            localCount := localCount + 1;
        ELSE
            status := WORD#16#8002;
        END_IF;
    END_IF;

    IF localRisingDequeue THEN
        IF localCount > 0 THEN
            item := buffer[localHead];
            localNext := localHead - localLower + 1;
            IF localNext >= localCapacity THEN
                localNext := 0;
            END_IF;
            localHead := localLower + localNext;
            localCount := localCount - 1;
        ELSE
            status := WORD#16#8001;
        END_IF;
    END_IF;
END_IF;

elementCount := localCount;

localLastEnqueue := enqueue;
localLastDequeue := dequeue;

END_FUNCTION_BLOCK

(* ---- public-medium-01.candidate_01.st ---- *)
TYPE ST_Pump :
STRUCT
    priority : INT;
    selection : BOOL;
    RunComd : BOOL;
END_STRUCT
END_TYPE;

FUNCTION_BLOCK FB_MultiPumpSwitchingControl
(* ENGINEERING_CONTRACT
   - mode=FALSE: manual mode; RunComd follows selection (PUB001/PUB002).
   - mode=TRUE: automatic mode; select three pumps with highest priority (PUB001/PUB003).
   - start: activates run enable; stop: deactivates run enable and stops all pumps (PUB002/PUB004).
   - Same-scan stop priority: if stop=TRUE, stop wins over start.
   - Run command is evaluated as selected AND run enable each scan.
   - Larger priority wins. Equal priority is unspecified; lower array index wins.
   - Mode transition with run enable retained is unspecified; retained run enable is used.
*)
(* CONTRACT_RULES [] *)
VAR
    runEnable : BOOL := FALSE;
    tmp_rank : INT;
    tmp_selected : ARRAY[1..5] OF BOOL;
    i : INT;
    j : INT;
END_VAR

IF stop THEN
    runEnable := FALSE;
ELSIF start THEN
    runEnable := TRUE;
END_IF;

IF mode THEN
    FOR i := 1 TO 5 DO
        tmp_rank := 0;
        FOR j := 1 TO 5 DO
            IF (pumpGroup[j].priority > pumpGroup[i].priority)
               OR ((pumpGroup[j].priority = pumpGroup[i].priority) AND (j < i)) THEN
                tmp_rank := tmp_rank + 1;
            END_IF;
        END_FOR;

        IF tmp_rank < 3 THEN
            tmp_selected[i] := TRUE;
        ELSE
            tmp_selected[i] := FALSE;
        END_IF;
    END_FOR;
ELSE
    FOR i := 1 TO 5 DO
        tmp_selected[i] := pumpGroup[i].selection;
    END_FOR;
END_IF;

FOR i := 1 TO 5 DO
    pumpGroup[i].RunComd := tmp_selected[i] AND runEnable;
END_FOR;

END_FUNCTION_BLOCK

(* ---- public-medium-01.candidate_02.st ---- *)
TYPE ST_Pump :
STRUCT
    priority : INT;
    selection : BOOL;
    RunComd : BOOL;
END_STRUCT
END_TYPE;

FUNCTION_BLOCK FB_MultiPumpSwitchingControl
(* ENGINEERING_CONTRACT
   - mode=FALSE: manual mode; RunComd follows selection (PUB001/PUB002).
   - mode=TRUE: automatic mode; select three pumps with highest priority (PUB001/PUB003).
   - start: activates run enable; stop: deactivates run enable and stops all pumps (PUB002/PUB004).
   - Same-scan stop priority: if stop=TRUE, stop wins over start.
   - Run command is evaluated as selected AND run enable each scan.
   - Larger priority wins. Equal priority is unspecified; lower array index wins.
   - Mode transition with run enable retained is unspecified; retained run enable is used.
*)
(* CONTRACT_RULES [] *)
VAR_INPUT
    mode : BOOL;
    start : BOOL;
    stop : BOOL;
END_VAR
VAR_IN_OUT
    pumpGroup : ARRAY[1..5] OF ST_Pump;
END_VAR
VAR
    runEnable : BOOL := FALSE;
    tmp_rank : INT;
    tmp_selected : ARRAY[1..5] OF BOOL;
    i : INT;
    j : INT;
END_VAR

IF stop THEN
    runEnable := FALSE;
ELSIF start THEN
    runEnable := TRUE;
END_IF;

IF mode THEN
    FOR i := 1 TO 5 DO
        tmp_rank := 0;
        FOR j := 1 TO 5 DO
            IF (pumpGroup[j].priority > pumpGroup[i].priority)
               OR ((pumpGroup[j].priority = pumpGroup[i].priority) AND (j < i)) THEN
                tmp_rank := tmp_rank + 1;
            END_IF;
        END_FOR;

        IF tmp_rank < 3 THEN
            tmp_selected[i] := TRUE;
        ELSE
            tmp_selected[i] := FALSE;
        END_IF;
    END_FOR;
ELSE
    FOR i := 1 TO 5 DO
        tmp_selected[i] := pumpGroup[i].selection;
    END_FOR;
END_IF;

FOR i := 1 TO 5 DO
    pumpGroup[i].RunComd := tmp_selected[i] AND runEnable;
END_FOR;

END_FUNCTION_BLOCK

(* ---- public-medium-01.raw_candidate_01.st ---- *)
TYPE ST_Pump :
STRUCT
    priority : INT;
    selection : BOOL;
    RunComd : BOOL;
END_STRUCT
END_TYPE

FUNCTION_BLOCK FB_MultiPumpSwitchingControl
(* ENGINEERING_CONTRACT
   - mode=FALSE: manual mode; RunComd follows selection (PUB001/PUB002).
   - mode=TRUE: automatic mode; select three pumps with highest priority (PUB001/PUB003).
   - start: activates run enable; stop: deactivates run enable and stops all pumps (PUB002/PUB004).
   - Same-scan stop priority: if stop=TRUE, stop wins over start.
   - Run command is evaluated as selected AND run enable each scan.
   - Larger priority wins. Equal priority is unspecified; lower array index wins.
   - Mode transition with run enable retained is unspecified; retained run enable is used.
*)
(* CONTRACT_RULES [] *)
VAR
    runEnable : BOOL := FALSE;
    tmp_rank : INT;
    tmp_selected : ARRAY[1..5] OF BOOL;
    i : INT;
    j : INT;
END_VAR

IF stop THEN
    runEnable := FALSE;
ELSIF start THEN
    runEnable := TRUE;
END_IF;

IF mode THEN
    FOR i := 1 TO 5 DO
        tmp_rank := 0;
        FOR j := 1 TO 5 DO
            IF (pumpGroup[j].priority > pumpGroup[i].priority)
               OR ((pumpGroup[j].priority = pumpGroup[i].priority) AND (j < i)) THEN
                tmp_rank := tmp_rank + 1;
            END_IF;
        END_FOR;

        IF tmp_rank < 3 THEN
            tmp_selected[i] := TRUE;
        ELSE
            tmp_selected[i] := FALSE;
        END_IF;
    END_FOR;
ELSE
    FOR i := 1 TO 5 DO
        tmp_selected[i] := pumpGroup[i].selection;
    END_FOR;
END_IF;

FOR i := 1 TO 5 DO
    pumpGroup[i].RunComd := tmp_selected[i] AND runEnable;
END_FOR;

END_FUNCTION_BLOCK

(* ---- public-medium-01.raw_candidate_02.st ---- *)
TYPE ST_Pump :
STRUCT
    priority : INT;
    selection : BOOL;
    RunComd : BOOL;
END_STRUCT
END_TYPE;

FUNCTION_BLOCK FB_MultiPumpSwitchingControl
(* ENGINEERING_CONTRACT
   - mode=FALSE: manual mode; RunComd follows selection (PUB001/PUB002).
   - mode=TRUE: automatic mode; select three pumps with highest priority (PUB001/PUB003).
   - start: activates run enable; stop: deactivates run enable and stops all pumps (PUB002/PUB004).
   - Same-scan stop priority: if stop=TRUE, stop wins over start.
   - Run command is evaluated as selected AND run enable each scan.
   - Larger priority wins. Equal priority is unspecified; lower array index wins.
   - Mode transition with run enable retained is unspecified; retained run enable is used.
*)
(* CONTRACT_RULES [] *)
VAR_INPUT
    mode : BOOL;
    start : BOOL;
    stop : BOOL;
END_VAR
VAR_IN_OUT
    pumpGroup : ARRAY[1..5] OF ST_Pump;
END_VAR
VAR
    runEnable : BOOL := FALSE;
    tmp_rank : INT;
    tmp_selected : ARRAY[1..5] OF BOOL;
    i : INT;
    j : INT;
END_VAR

IF stop THEN
    runEnable := FALSE;
ELSIF start THEN
    runEnable := TRUE;
END_IF;

IF mode THEN
    FOR i := 1 TO 5 DO
        tmp_rank := 0;
        FOR j := 1 TO 5 DO
            IF (pumpGroup[j].priority > pumpGroup[i].priority)
               OR ((pumpGroup[j].priority = pumpGroup[i].priority) AND (j < i)) THEN
                tmp_rank := tmp_rank + 1;
            END_IF;
        END_FOR;

        IF tmp_rank < 3 THEN
            tmp_selected[i] := TRUE;
        ELSE
            tmp_selected[i] := FALSE;
        END_IF;
    END_FOR;
ELSE
    FOR i := 1 TO 5 DO
        tmp_selected[i] := pumpGroup[i].selection;
    END_FOR;
END_IF;

FOR i := 1 TO 5 DO
    pumpGroup[i].RunComd := tmp_selected[i] AND runEnable;
END_FOR;

END_FUNCTION_BLOCK

(* ---- public-medium-02.candidate_01.st ---- *)
TYPE ST_AnalogChannel :
STRUCT
    enable : BOOL;
    hiLIM : REAL;
    loLIM : REAL;
    bipolar : BOOL;
    measuringMode : INT;
    retVal : WORD;
    outputValue : REAL;
END_STRUCT
END_TYPE;

(* ENGINEERING_CONTRACT
   count: process ordinal positions 0..count-1 from each array's own lower bound, limited to both upper bounds.
   enable=FALSE: channel is skipped; retVal/outputValue are not written (unspecified by PUB002).
   mode invalid: retVal=16#8001, outputValue unchanged, conversion skipped (PUB006).
   hiLIM<=loLIM: retVal=16#8002, outputValue unchanged, conversion skipped (PUB007).
   success: retVal=16#0000, outputValue set from analogValues[ordinal] (PUB003/PUB004/PUB005).
   mode0 unipolar: loLIM + raw/27648*(hiLIM-loLIM); bipolar: loLIM + (raw+27648)/55296*(hiLIM-loLIM).
   mode1: raw/10.0; mode2: raw/100.0. Raw INT converted explicitly to REAL.
   no latches/edges/retention; each invocation recomputes selected enabled channels (PUB001).
*)

(* CONTRACT_RULES [] *)

FUNCTION_BLOCK AnalogBatchProcessing
VAR_INPUT
    count : DINT;
END_VAR
VAR_IN_OUT
    analogValues : ARRAY[*] OF INT;
    channels : ARRAY[*] OF ST_AnalogChannel;
END_VAR
VAR
    tmp_i : DINT;
    tmp_process_count : DINT;
    tmp_analog_lower : DINT;
    tmp_channel_lower : DINT;
    tmp_analog_len : DINT;
    tmp_channel_len : DINT;
    tmp_analog_index : DINT;
    tmp_channel_index : DINT;
    tmp_raw : REAL;
END_VAR

tmp_analog_lower := LOWER_BOUND(analogValues, 1);
tmp_channel_lower := LOWER_BOUND(channels, 1);
tmp_analog_len := UPPER_BOUND(analogValues, 1) - tmp_analog_lower + 1;
tmp_channel_len := UPPER_BOUND(channels, 1) - tmp_channel_lower + 1;

tmp_process_count := count;
IF tmp_process_count < 0 THEN
    tmp_process_count := 0;
END_IF;
IF tmp_process_count > tmp_analog_len THEN
    tmp_process_count := tmp_analog_len;
END_IF;
IF tmp_process_count > tmp_channel_len THEN
    tmp_process_count := tmp_channel_len;
END_IF;

FOR tmp_i := 0 TO tmp_process_count - 1 DO
    tmp_analog_index := tmp_analog_lower + tmp_i;
    tmp_channel_index := tmp_channel_lower + tmp_i;

    IF channels[tmp_channel_index].enable THEN
        IF (channels[tmp_channel_index].measuringMode <> 0)
           AND (channels[tmp_channel_index].measuringMode <> 1)
           AND (channels[tmp_channel_index].measuringMode <> 2) THEN
            channels[tmp_channel_index].retVal := 16#8001;
        ELSIF channels[tmp_channel_index].hiLIM <= channels[tmp_channel_index].loLIM THEN
            channels[tmp_channel_index].retVal := 16#8002;
        ELSE
            tmp_raw := INT_TO_REAL(analogValues[tmp_analog_index]);

            CASE channels[tmp_channel_index].measuringMode OF
                0:
                    IF channels[tmp_channel_index].bipolar THEN
                        channels[tmp_channel_index].outputValue :=
                            channels[tmp_channel_index].loLIM
                            + ((tmp_raw + 27648.0) / 55296.0)
                            * (channels[tmp_channel_index].hiLIM - channels[tmp_channel_index].loLIM);
                    ELSE
                        channels[tmp_channel_index].outputValue :=
                            channels[tmp_channel_index].loLIM
                            + (tmp_raw / 27648.0)
                            * (channels[tmp_channel_index].hiLIM - channels[tmp_channel_index].loLIM);
                    END_IF;
                1:
                    channels[tmp_channel_index].outputValue := tmp_raw / 10.0;
                2:
                    channels[tmp_channel_index].outputValue := tmp_raw / 100.0;
            END_CASE;

            channels[tmp_channel_index].retVal := 16#0000;
        END_IF;
    END_IF;
END_FOR;

END_FUNCTION_BLOCK

(* ---- public-medium-02.raw_candidate_01.st ---- *)
TYPE ST_AnalogChannel :
STRUCT
    enable : BOOL;
    hiLIM : REAL;
    loLIM : REAL;
    bipolar : BOOL;
    measuringMode : INT;
    retVal : WORD;
    outputValue : REAL;
END_STRUCT
END_TYPE

(* ENGINEERING_CONTRACT
   count: process ordinal positions 0..count-1 from each array's own lower bound, limited to both upper bounds.
   enable=FALSE: channel is skipped; retVal/outputValue are not written (unspecified by PUB002).
   mode invalid: retVal=16#8001, outputValue unchanged, conversion skipped (PUB006).
   hiLIM<=loLIM: retVal=16#8002, outputValue unchanged, conversion skipped (PUB007).
   success: retVal=16#0000, outputValue set from analogValues[ordinal] (PUB003/PUB004/PUB005).
   mode0 unipolar: loLIM + raw/27648*(hiLIM-loLIM); bipolar: loLIM + (raw+27648)/55296*(hiLIM-loLIM).
   mode1: raw/10.0; mode2: raw/100.0. Raw INT converted explicitly to REAL.
   no latches/edges/retention; each invocation recomputes selected enabled channels (PUB001).
*)

(* CONTRACT_RULES [] *)

FUNCTION_BLOCK AnalogBatchProcessing
VAR_INPUT
    count : DINT;
END_VAR
VAR_IN_OUT
    analogValues : ARRAY[*] OF INT;
    channels : ARRAY[*] OF ST_AnalogChannel;
END_VAR
VAR
    tmp_i : DINT;
    tmp_process_count : DINT;
    tmp_analog_lower : DINT;
    tmp_channel_lower : DINT;
    tmp_analog_len : DINT;
    tmp_channel_len : DINT;
    tmp_analog_index : DINT;
    tmp_channel_index : DINT;
    tmp_raw : REAL;
END_VAR

tmp_analog_lower := LOWER_BOUND(analogValues, 1);
tmp_channel_lower := LOWER_BOUND(channels, 1);
tmp_analog_len := UPPER_BOUND(analogValues, 1) - tmp_analog_lower + 1;
tmp_channel_len := UPPER_BOUND(channels, 1) - tmp_channel_lower + 1;

tmp_process_count := count;
IF tmp_process_count < 0 THEN
    tmp_process_count := 0;
END_IF;
IF tmp_process_count > tmp_analog_len THEN
    tmp_process_count := tmp_analog_len;
END_IF;
IF tmp_process_count > tmp_channel_len THEN
    tmp_process_count := tmp_channel_len;
END_IF;

FOR tmp_i := 0 TO tmp_process_count - 1 DO
    tmp_analog_index := tmp_analog_lower + tmp_i;
    tmp_channel_index := tmp_channel_lower + tmp_i;

    IF channels[tmp_channel_index].enable THEN
        IF (channels[tmp_channel_index].measuringMode <> 0)
           AND (channels[tmp_channel_index].measuringMode <> 1)
           AND (channels[tmp_channel_index].measuringMode <> 2) THEN
            channels[tmp_channel_index].retVal := 16#8001;
        ELSIF channels[tmp_channel_index].hiLIM <= channels[tmp_channel_index].loLIM THEN
            channels[tmp_channel_index].retVal := 16#8002;
        ELSE
            tmp_raw := INT_TO_REAL(analogValues[tmp_analog_index]);

            CASE channels[tmp_channel_index].measuringMode OF
                0:
                    IF channels[tmp_channel_index].bipolar THEN
                        channels[tmp_channel_index].outputValue :=
                            channels[tmp_channel_index].loLIM
                            + ((tmp_raw + 27648.0) / 55296.0)
                            * (channels[tmp_channel_index].hiLIM - channels[tmp_channel_index].loLIM);
                    ELSE
                        channels[tmp_channel_index].outputValue :=
                            channels[tmp_channel_index].loLIM
                            + (tmp_raw / 27648.0)
                            * (channels[tmp_channel_index].hiLIM - channels[tmp_channel_index].loLIM);
                    END_IF;
                1:
                    channels[tmp_channel_index].outputValue := tmp_raw / 10.0;
                2:
                    channels[tmp_channel_index].outputValue := tmp_raw / 100.0;
            END_CASE;

            channels[tmp_channel_index].retVal := 16#0000;
        END_IF;
    END_IF;
END_FOR;

END_FUNCTION_BLOCK

(* ---- public-medium-03.candidate_01.st ---- *)
FUNCTION_BLOCK FB
VAR_INPUT
    cyclicExecution : BOOL;
    trigger : BOOL;
    value : LREAL;
    windowSize : INT;
    reset : BOOL;
END_VAR
VAR_OUTPUT
    average : LREAL;
    windowSizeReached : BOOL;
    error : BOOL;
    status : WORD;
END_VAR
VAR
    local_triggerEdge : R_TRIG;
    local_samples : ARRAY[0..99] OF LREAL;
    local_sampleCount : INT;
    local_index : INT;
    local_limit : INT;
    local_sum : LREAL;
END_VAR

(*
ENGINEERING_CONTRACT
average: activation = each valid acquisition (cyclicExecution TRUE every scan, or trigger rising edge while cyclicExecution FALSE); retention = holds last computed value until next acquisition; explicit reset = reset TRUE; same-scan priority = reset before acquisition; invalid window also clears calculation state in this implementation; units LREAL.
windowSizeReached: activation = sampleCount >= valid windowSize; retention = remains TRUE once reached; explicit reset = reset TRUE; invalid window clears it.
error/status: error FALSE + status 16#0000 on valid window; error TRUE + status 16#8200 when windowSize < 1 or windowSize > 100; invalid window is checked first.
trigger/cyclic: cyclicExecution TRUE disables trigger; trigger uses rising edge only. PUB001-PUB007.
*)

(* CONTRACT_RULES [] *)

local_triggerEdge(CLK := trigger);

error := FALSE;
status := 16#0000;

IF (windowSize < 1) OR (windowSize > 100) THEN
    error := TRUE;
    status := 16#8200;
    average := 0.0;
    windowSizeReached := FALSE;
    local_sampleCount := 0;
    RETURN;
END_IF;

IF local_sampleCount >= windowSize THEN
    windowSizeReached := TRUE;
ELSE
    windowSizeReached := FALSE;
END_IF;

IF reset THEN
    local_sampleCount := 0;
    average := 0.0;
    windowSizeReached := FALSE;
    RETURN;
END_IF;

IF cyclicExecution OR local_triggerEdge.Q THEN
    IF local_sampleCount < 100 THEN
        local_sampleCount := local_sampleCount + 1;
    END_IF;

    FOR local_index := 99 TO 1 BY -1 DO
        local_samples[local_index] := local_samples[local_index - 1];
    END_FOR;
    local_samples[0] := value;

    local_limit := windowSize;
    IF local_limit > local_sampleCount THEN
        local_limit := local_sampleCount;
    END_IF;

    local_sum := 0.0;
    IF local_limit > 0 THEN
        FOR local_index := 0 TO local_limit - 1 DO
            local_sum := local_sum + local_samples[local_index];
        END_FOR;
        average := local_sum / INT_TO_LREAL(local_limit);
    ELSE
        average := 0.0;
    END_IF;

    IF local_sampleCount >= windowSize THEN
        windowSizeReached := TRUE;
    ELSE
        windowSizeReached := FALSE;
    END_IF;
END_IF;

END_FUNCTION_BLOCK

(* ---- public-medium-03.raw_candidate_01.st ---- *)
FUNCTION_BLOCK FB
VAR_INPUT
    cyclicExecution : BOOL;
    trigger : BOOL;
    value : LREAL;
    windowSize : INT;
    reset : BOOL;
END_VAR
VAR_OUTPUT
    average : LREAL;
    windowSizeReached : BOOL;
    error : BOOL;
    status : WORD;
END_VAR
VAR
    local_triggerEdge : R_TRIG;
    local_samples : ARRAY[0..99] OF LREAL;
    local_sampleCount : INT;
    local_index : INT;
    local_limit : INT;
    local_sum : LREAL;
END_VAR

(*
ENGINEERING_CONTRACT
average: activation = each valid acquisition (cyclicExecution TRUE every scan, or trigger rising edge while cyclicExecution FALSE); retention = holds last computed value until next acquisition; explicit reset = reset TRUE; same-scan priority = reset before acquisition; invalid window also clears calculation state in this implementation; units LREAL.
windowSizeReached: activation = sampleCount >= valid windowSize; retention = remains TRUE once reached; explicit reset = reset TRUE; invalid window clears it.
error/status: error FALSE + status 16#0000 on valid window; error TRUE + status 16#8200 when windowSize < 1 or windowSize > 100; invalid window is checked first.
trigger/cyclic: cyclicExecution TRUE disables trigger; trigger uses rising edge only. PUB001-PUB007.
*)

(* CONTRACT_RULES [] *)

local_triggerEdge(CLK := trigger);

error := FALSE;
status := 16#0000;

IF (windowSize < 1) OR (windowSize > 100) THEN
    error := TRUE;
    status := 16#8200;
    average := 0.0;
    windowSizeReached := FALSE;
    local_sampleCount := 0;
    RETURN;
END_IF;

IF local_sampleCount >= windowSize THEN
    windowSizeReached := TRUE;
ELSE
    windowSizeReached := FALSE;
END_IF;

IF reset THEN
    local_sampleCount := 0;
    average := 0.0;
    windowSizeReached := FALSE;
    RETURN;
END_IF;

IF cyclicExecution OR local_triggerEdge.Q THEN
    IF local_sampleCount < 100 THEN
        local_sampleCount := local_sampleCount + 1;
    END_IF;

    FOR local_index := 99 TO 1 BY -1 DO
        local_samples[local_index] := local_samples[local_index - 1];
    END_FOR;
    local_samples[0] := value;

    local_limit := windowSize;
    IF local_limit > local_sampleCount THEN
        local_limit := local_sampleCount;
    END_IF;

    local_sum := 0.0;
    IF local_limit > 0 THEN
        FOR local_index := 0 TO local_limit - 1 DO
            local_sum := local_sum + local_samples[local_index];
        END_FOR;
        average := local_sum / INT_TO_LREAL(local_limit);
    ELSE
        average := 0.0;
    END_IF;

    IF local_sampleCount >= windowSize THEN
        windowSizeReached := TRUE;
    ELSE
        windowSizeReached := FALSE;
    END_IF;
END_IF;

END_FUNCTION_BLOCK

(* ---- public-medium-04.candidate_01.st ---- *)
(* ENGINEERING_CONTRACT
- CurrentTemperature: unconditional pass-through each scan; no hold/reset; temperature units are unspecified.
- SetTempDisplay: unconditional pass-through each scan; no hold/reset; temperature units are unspecified.
- HeaterStatus: mirrors HeaterOutput every scan; no hold/reset.
- HeaterOutput: active when sensor is valid and temperature < setpoint and no overheat; off on >=, fault, or overheat; no latch. PUB003/PUB004/PUB007.
- OverheatProtection: set after heater runs continuously >5000 ms; held for at least 3000 ms, then auto-clears; no manual reset. PUB005.
- Same-scan priority: sensor fault and active overheat force heater off; after the 3s wait elapses, normal heater control can resume in the same scan.
- Boundaries: sensor fault is <0.0 or >100.0; strict >5s uses T#5001MS; cool-down wait uses T#3S.
*)
(* CONTRACT_RULES [] *)

FUNCTION_BLOCK FB
VAR_INPUT
    TemperatureSensorInput : REAL;
    SetTemperature : REAL;
END_VAR

VAR_OUTPUT
    CurrentTemperature : REAL;
    SetTempDisplay : REAL;
    HeaterStatus : BOOL;
    OverheatProtection : BOOL;
    HeaterOutput : BOOL;
END_VAR

VAR
    local_SensorFault : BOOL;
    local_BaseHeaterRequest : BOOL;
    local_HeaterAllowed : BOOL;
    local_OverheatActive : BOOL;
    local_HeaterRunTimer : TON;
    local_CooldownTimer : TON;
END_VAR

local_SensorFault := (TemperatureSensorInput < 0.0) OR (TemperatureSensorInput > 100.0);
local_BaseHeaterRequest := (NOT local_SensorFault) AND (TemperatureSensorInput < SetTemperature);

IF local_OverheatActive THEN
    local_CooldownTimer(IN := TRUE, PT := T#3S);
    local_HeaterAllowed := FALSE;

    IF local_CooldownTimer.Q THEN
        local_OverheatActive := FALSE;
        local_HeaterAllowed := local_BaseHeaterRequest;
    END_IF;

    local_HeaterRunTimer(IN := local_HeaterAllowed, PT := T#5001MS);

    IF local_HeaterRunTimer.Q THEN
        local_OverheatActive := TRUE;
        local_HeaterAllowed := FALSE;
    END_IF;
ELSE
    local_CooldownTimer(IN := FALSE, PT := T#3S);
    local_HeaterAllowed := local_BaseHeaterRequest;

    local_HeaterRunTimer(IN := local_HeaterAllowed, PT := T#5001MS);

    IF local_HeaterRunTimer.Q THEN
        local_OverheatActive := TRUE;
        local_HeaterAllowed := FALSE;
    END_IF;
END_IF;

HeaterOutput := (NOT local_SensorFault) AND local_HeaterAllowed;
HeaterStatus := HeaterOutput;
OverheatProtection := local_OverheatActive;
CurrentTemperature := TemperatureSensorInput;
SetTempDisplay := SetTemperature;

END_FUNCTION_BLOCK

(* ---- public-medium-04.raw_candidate_01.st ---- *)
(* ENGINEERING_CONTRACT
- CurrentTemperature: unconditional pass-through each scan; no hold/reset; temperature units are unspecified.
- SetTempDisplay: unconditional pass-through each scan; no hold/reset; temperature units are unspecified.
- HeaterStatus: mirrors HeaterOutput every scan; no hold/reset.
- HeaterOutput: active when sensor is valid and temperature < setpoint and no overheat; off on >=, fault, or overheat; no latch. PUB003/PUB004/PUB007.
- OverheatProtection: set after heater runs continuously >5000 ms; held for at least 3000 ms, then auto-clears; no manual reset. PUB005.
- Same-scan priority: sensor fault and active overheat force heater off; after the 3s wait elapses, normal heater control can resume in the same scan.
- Boundaries: sensor fault is <0.0 or >100.0; strict >5s uses T#5001MS; cool-down wait uses T#3S.
*)
(* CONTRACT_RULES [] *)

FUNCTION_BLOCK FB
VAR_INPUT
    TemperatureSensorInput : REAL;
    SetTemperature : REAL;
END_VAR

VAR_OUTPUT
    CurrentTemperature : REAL;
    SetTempDisplay : REAL;
    HeaterStatus : BOOL;
    OverheatProtection : BOOL;
    HeaterOutput : BOOL;
END_VAR

VAR
    local_SensorFault : BOOL;
    local_BaseHeaterRequest : BOOL;
    local_HeaterAllowed : BOOL;
    local_OverheatActive : BOOL;
    local_HeaterRunTimer : TON;
    local_CooldownTimer : TON;
END_VAR

local_SensorFault := (TemperatureSensorInput < 0.0) OR (TemperatureSensorInput > 100.0);
local_BaseHeaterRequest := (NOT local_SensorFault) AND (TemperatureSensorInput < SetTemperature);

IF local_OverheatActive THEN
    local_CooldownTimer(IN := TRUE, PT := T#3S);
    local_HeaterAllowed := FALSE;

    IF local_CooldownTimer.Q THEN
        local_OverheatActive := FALSE;
        local_HeaterAllowed := local_BaseHeaterRequest;
    END_IF;

    local_HeaterRunTimer(IN := local_HeaterAllowed, PT := T#5001MS);

    IF local_HeaterRunTimer.Q THEN
        local_OverheatActive := TRUE;
        local_HeaterAllowed := FALSE;
    END_IF;
ELSE
    local_CooldownTimer(IN := FALSE, PT := T#3S);
    local_HeaterAllowed := local_BaseHeaterRequest;

    local_HeaterRunTimer(IN := local_HeaterAllowed, PT := T#5001MS);

    IF local_HeaterRunTimer.Q THEN
        local_OverheatActive := TRUE;
        local_HeaterAllowed := FALSE;
    END_IF;
END_IF;

HeaterOutput := (NOT local_SensorFault) AND local_HeaterAllowed;
HeaterStatus := HeaterOutput;
OverheatProtection := local_OverheatActive;
CurrentTemperature := TemperatureSensorInput;
SetTempDisplay := SetTemperature;

END_FUNCTION_BLOCK

(* ---- public-medium-05.candidate_01.st ---- *)
FUNCTION_BLOCK ProductionLineControl
(*
ENGINEERING_CONTRACT
MotorForward (PUB001/PUB002/PUB003): activate manual ForwardButton or auto transfer state; hold through transfer to destination sensor; deactivate at destination sensor, manual release, or not in transfer state; simultaneous manual Forward/Reverse is interlocked, no motion.
MotorReverse (PUB002): activate only manual ReverseButton; no hold; deactivate on release or ForwardButton.
CompletionLight (PUB003): activate in auto at C while SensorC and ButtonC are TRUE; retain while SensorC remains TRUE; deactivation only when SensorC becomes FALSE; manual Mode does not reset it.
Bounds/units: BOOL inputs, BOOL outputs, discrete scan steps; buttons are level-gated, not edge-only.
Unspecified: simultaneous manual Forward/Reverse means no motion; automatic step is retained across mode changes.
*)
(* CONTRACT_RULES [] *)
VAR_INPUT
    Mode : BOOL;
    ForwardButton : BOOL;
    ReverseButton : BOOL;
    SensorA : BOOL;
    SensorB : BOOL;
    SensorC : BOOL;
    ButtonA : BOOL;
    ButtonB : BOOL;
    ButtonC : BOOL;
END_VAR
VAR_OUTPUT
    MotorForward : BOOL;
    MotorReverse : BOOL;
    CompletionLight : BOOL;
END_VAR
VAR
    AutoStep : INT := 0;
END_VAR

MotorForward := FALSE;
MotorReverse := FALSE;

IF NOT SensorC THEN
    CompletionLight := FALSE;
END_IF;

IF Mode THEN
    CASE AutoStep OF
        0:
            IF SensorA AND ButtonA THEN
                AutoStep := 1;
                MotorForward := TRUE;
            END_IF;

        1:
            IF SensorB THEN
                AutoStep := 2;
            END_IF;

        2:
            IF ButtonB THEN
                AutoStep := 3;
                MotorForward := TRUE;
            END_IF;

        3:
            IF SensorC THEN
                AutoStep := 4;
            END_IF;

        4:
            IF SensorC AND ButtonC THEN
                CompletionLight := TRUE;
            END_IF;
            IF NOT SensorC THEN
                AutoStep := 0;
            END_IF;
    END_CASE;
ELSE
    MotorForward := ForwardButton AND NOT ReverseButton;
    MotorReverse := ReverseButton AND NOT ForwardButton;
END_IF;
END_FUNCTION_BLOCK
